DATA_BLOCK DB 1
VERSION : 0.1


  STRUCT
   STAT0 : CHAR ;
   STAT1 : CHAR ;
   STAT2 : CHAR ;
   STAT3 : CHAR ;
   STAT4 : CHAR ;
   STAT5 : CHAR ;
   STAT6 : CHAR ;
   STAT7 : CHAR ;
   STAT8 : CHAR ;
   STAT9 : CHAR ;
   STAT10 : CHAR ;
   STAT11 : CHAR ;
  END_STRUCT ;
BEGIN
   STAT0 := ' ';
   STAT1 := ' ';
   STAT2 := ' ';
   STAT3 := ' ';
   STAT4 := ' ';
   STAT5 := ' ';
   STAT6 := ' ';
   STAT7 := ' ';
   STAT8 := ' ';
   STAT9 := ' ';
   STAT10 := ' ';
   STAT11 := ' ';
END_DATA_BLOCK

DATA_BLOCK DB 2
VERSION : 0.1


  STRUCT
   STAT0 : CHAR ;
   STAT1 : CHAR ;
   STAT2 : CHAR ;
   STAT3 : CHAR ;
   STAT4 : CHAR ;
   STAT5 : CHAR ;
   STAT6 : CHAR ;
   STAT7 : CHAR ;
  END_STRUCT ;
BEGIN
   STAT0 := ' ';
   STAT1 := ' ';
   STAT2 := ' ';
   STAT3 := ' ';
   STAT4 := ' ';
   STAT5 := ' ';
   STAT6 := ' ';
   STAT7 := ' ';
END_DATA_BLOCK

DATA_BLOCK DB 3
VERSION : 0.1


  STRUCT
   STAT0 : INT ;
   STAT1 : BOOL ;
   STAT2 : INT ;
   STAT3 : BOOL ;
   STAT4 : BOOL ;
   STAT5 : BOOL ;
   STAT6 : BOOL ;
   STAT7 : BOOL ;
   STAT8 : BOOL ;
   STAT9 : BOOL ;
   STAT10 : BOOL ;
   STAT11 : BOOL ;
   STAT12 : BOOL ;
   STAT13 : BOOL ;
   STAT14 : BOOL ;
   STAT15 : INT ;
   STAT16 : INT ;
   STAT17 : INT ;
   STAT18 : INT ;
   STAT19 : CHAR  := '2';
   STAT20 : CHAR  := '8';
   STAT21 : INT ;
   STAT22 : CHAR  := '-';
   STAT23 : CHAR  := '-';
   STAT24 : CHAR  := '-';
   STAT25 : CHAR  := '-';
   STAT26 : CHAR  := '-';
   STAT27 : CHAR  := '-';
   STAT28 : CHAR  := '-';
   STAT29 : CHAR  := '-';
   STAT30 : CHAR  := '-';
   STAT31 : CHAR  := '-';
   STAT32 : CHAR  := '-';
   STAT33 : CHAR  := '-';
   STAT34 : CHAR  := '-';
   STAT35 : CHAR  := '-';
   STAT36 : CHAR  := '-';
   STAT37 : CHAR  := '-';
   STAT38 : CHAR  := '-';
   STAT39 : CHAR  := '-';
   STAT40 : CHAR  := '1';
   STAT41 : CHAR  := '2';
   STAT42 : CHAR  := '3';
   STAT43 : CHAR  := '4';
   STAT44 : CHAR  := '5';
   STAT45 : CHAR  := '6';
   STAT46 : CHAR  := '7';
   STAT47 : CHAR  := '8';
   STAT48 : CHAR  := '9';
   STAT49 : CHAR  := '0';
   STAT50 : INT ;
   STAT51 : INT ;
   STAT52 : INT ;
   STAT53 : INT ;
   STAT54 : INT ;
   STAT55 : CHAR  := '1';
   STAT56 : CHAR  := '4';
   STAT57 : CHAR  := '6';
   STAT58 : CHAR  := '1';
   STAT59 : CHAR  := '2';
   STAT60 : CHAR  := '3';
   STAT61 : CHAR  := '4';
   STAT62 : CHAR  := '5';
   STAT63 : CHAR  := '6';
   STAT64 : CHAR  := '7';
   STAT65 : CHAR  := '8';
   STAT66 : CHAR  := '9';
   STAT67 : CHAR  := '0';
   STAT68 : CHAR  := '1';
   STAT69 : CHAR  := '2';
   STAT70 : CHAR  := '3';
   STAT71 : CHAR  := '4';
   STAT72 : CHAR  := '5';
   STAT73 : CHAR  := '6';
   STAT74 : CHAR  := '7';
   STAT75 : CHAR  := '8';
   STAT76 : CHAR  := 'P';
   STAT77 : CHAR  := 'P';
   STAT78 : CHAR  := 'P';
   STAT79 : INT ;
   STAT80 : CHAR  := '0';
   STAT81 : CHAR  := '0';
   STAT82 : CHAR  := '0';
   STAT83 : CHAR  := '0';
   STAT84 : CHAR  := '0';
   STAT85 : CHAR  := '0';
   STAT86 : INT ;
   STAT87 : CHAR ;
   STAT88 : INT ;
   STAT89 : BOOL ;
   STAT90 : BOOL ;
   STAT91 : CHAR ;
   STAT92 : CHAR ;
   STAT93 : CHAR ;
   STAT94 : CHAR ;
   STAT95 : CHAR ;
   STAT96 : CHAR ;
   STAT97 : CHAR ;
   STAT98 : CHAR ;
   STAT99 : CHAR ;
   STAT100 : CHAR ;
   STAT101 : CHAR ;
   STAT102 : CHAR ;
   STAT103 : ARRAY  [1 .. 3 ] OF CHAR ;
   STAT104 : BOOL ;
   STAT105 : ARRAY  [1 .. 10 ] OF STRUCT
    STAT106 : REAL ;
    STAT107 : REAL ;
    STAT108 : REAL ;
   END_STRUCT ;
   STAT109 : CHAR ;
   STAT110 : CHAR ;
   STAT111 : ARRAY  [1 .. 10 ] OF REAL ;
   STAT112 : INT ;
   STAT113 : BOOL ;
   STAT114 : BOOL ;
   STAT115 : BOOL ;
  END_STRUCT ;
BEGIN
   STAT0 := 0;
   STAT1 := FALSE;
   STAT2 := 0;
   STAT3 := FALSE;
   STAT4 := FALSE;
   STAT5 := FALSE;
   STAT6 := FALSE;
   STAT7 := FALSE;
   STAT8 := FALSE;
   STAT9 := FALSE;
   STAT10 := FALSE;
   STAT11 := FALSE;
   STAT12 := FALSE;
   STAT13 := FALSE;
   STAT14 := FALSE;
   STAT15 := 0;
   STAT16 := 0;
   STAT17 := 0;
   STAT18 := 0;
   STAT19 := ' ';
   STAT20 := ' ';
   STAT21 := 0;
   STAT22 := '1';
   STAT23 := '2';
   STAT24 := '3';
   STAT25 := '4';
   STAT26 := '5';
   STAT27 := '$00';
   STAT28 := '7';
   STAT29 := '8';
   STAT30 := '9';
   STAT31 := '0';
   STAT32 := '1';
   STAT33 := '$00';
   STAT34 := '3';
   STAT35 := '4';
   STAT36 := '5';
   STAT37 := '6';
   STAT38 := '7';
   STAT39 := '$00';
   STAT40 := '-';
   STAT41 := '-';
   STAT42 := '-';
   STAT43 := '-';
   STAT44 := '-';
   STAT45 := '-';
   STAT46 := '-';
   STAT47 := '-';
   STAT48 := '-';
   STAT49 := '-';
   STAT50 := 0;
   STAT51 := 0;
   STAT52 := 0;
   STAT53 := 0;
   STAT54 := 0;
   STAT55 := '1';
   STAT56 := '2';
   STAT57 := '3';
   STAT58 := '$00';
   STAT59 := '$00';
   STAT60 := '$00';
   STAT61 := '$00';
   STAT62 := '$00';
   STAT63 := '$00';
   STAT64 := '$00';
   STAT65 := '$00';
   STAT66 := '$00';
   STAT67 := '$00';
   STAT68 := '$00';
   STAT69 := '$00';
   STAT70 := '$00';
   STAT71 := '$00';
   STAT72 := '$00';
   STAT73 := '$00';
   STAT74 := '$00';
   STAT75 := '$00';
   STAT76 := 'P';
   STAT77 := 'P';
   STAT78 := 'P';
   STAT79 := 0;
   STAT80 := '$00';
   STAT81 := '$00';
   STAT82 := '$00';
   STAT83 := '$00';
   STAT84 := '$00';
   STAT85 := '$00';
   STAT86 := 1;
   STAT87 := '1';
   STAT88 := 49;
   STAT89 := FALSE;
   STAT90 := FALSE;
   STAT91 := '-';
   STAT92 := '-';
   STAT93 := '-';
   STAT94 := '$00';
   STAT95 := '$00';
   STAT96 := '$00';
   STAT97 := '$00';
   STAT98 := '$00';
   STAT99 := '$00';
   STAT100 := '$00';
   STAT101 := '$00';
   STAT102 := '$00';
   STAT103[1] := '-';
   STAT103[2] := '-';
   STAT103[3] := '-';
   STAT104 := FALSE;
   STAT105[1].STAT106 := 1.616663e+004;
   STAT105[1].STAT107 := -7.696248e+003;
   STAT105[1].STAT108 := 1.325872e+004;
   STAT105[2].STAT106 := -8.515102e+003;
   STAT105[2].STAT107 := 3.194731e+000;
   STAT105[2].STAT108 := 2.146098e+004;
   STAT105[3].STAT106 := -3.152269e+003;
   STAT105[3].STAT107 := 5.230335e+001;
   STAT105[3].STAT108 := 1.702762e+004;
   STAT105[4].STAT106 := 4.876809e+003;
   STAT105[4].STAT107 := -1.412248e+003;
   STAT105[4].STAT108 := 3.514912e+004;
   STAT105[5].STAT106 := 0.000000e+000;
   STAT105[5].STAT107 := 0.000000e+000;
   STAT105[5].STAT108 := 0.000000e+000;
   STAT105[6].STAT106 := 0.000000e+000;
   STAT105[6].STAT107 := 0.000000e+000;
   STAT105[6].STAT108 := 0.000000e+000;
   STAT105[7].STAT106 := 0.000000e+000;
   STAT105[7].STAT107 := 0.000000e+000;
   STAT105[7].STAT108 := 0.000000e+000;
   STAT105[8].STAT106 := 0.000000e+000;
   STAT105[8].STAT107 := 0.000000e+000;
   STAT105[8].STAT108 := 0.000000e+000;
   STAT105[9].STAT106 := 0.000000e+000;
   STAT105[9].STAT107 := 0.000000e+000;
   STAT105[9].STAT108 := 0.000000e+000;
   STAT105[10].STAT106 := 0.000000e+000;
   STAT105[10].STAT107 := 0.000000e+000;
   STAT105[10].STAT108 := 0.000000e+000;
   STAT109 := '-';
   STAT110 := '-';
   STAT111[1] := -2.054582e+003;
   STAT111[2] := -2.149658e-001;
   STAT111[3] := -9.505859e+000;
   STAT111[4] := 1.638507e+003;
   STAT111[5] := 0.000000e+000;
   STAT111[6] := 0.000000e+000;
   STAT111[7] := 0.000000e+000;
   STAT111[8] := 0.000000e+000;
   STAT111[9] := 0.000000e+000;
   STAT111[10] := 0.000000e+000;
   STAT112 := 1;
   STAT113 := FALSE;
   STAT114 := FALSE;
   STAT115 := FALSE;
END_DATA_BLOCK

DATA_BLOCK DB 4
VERSION : 0.1


  STRUCT
   STAT0 : INT ;
   STAT1 : ARRAY  [1 .. 10 ] OF INT ;
   STAT2 : ARRAY  [1 .. 10 ] OF INT ;
   STAT3 : ARRAY  [1 .. 10 ] OF INT ;
  END_STRUCT ;
BEGIN
   STAT0 := 0;
   STAT1[1] := -32768;
   STAT1[2] := 17072;
   STAT1[3] := 17056;
   STAT1[4] := 16968;
   STAT1[5] := 0;
   STAT1[6] := 0;
   STAT1[7] := 0;
   STAT1[8] := 0;
   STAT1[9] := 0;
   STAT1[10] := 0;
   STAT2[1] := 5576;
   STAT2[2] := 1968;
   STAT2[3] := -1312;
   STAT2[4] := -1624;
   STAT2[5] := 0;
   STAT2[6] := 0;
   STAT2[7] := 0;
   STAT2[8] := 0;
   STAT2[9] := 0;
   STAT2[10] := 0;
   STAT3[1] := -1632;
   STAT3[2] := 13768;
   STAT3[3] := 27488;
   STAT3[4] := 27496;
   STAT3[5] := 0;
   STAT3[6] := 0;
   STAT3[7] := 0;
   STAT3[8] := 0;
   STAT3[9] := 0;
   STAT3[10] := 0;
END_DATA_BLOCK

DATA_BLOCK DB 5
VERSION : 0.1


  STRUCT
   STAT0 : INT ;
   STAT1 : ARRAY  [1 .. 10 ] OF BOOL ;
   STAT2 : ARRAY  [1 .. 10 ] OF BOOL ;
   STAT3 : BOOL ;
   STAT4 : BOOL ;
   STAT5 : BOOL ;
   STAT6 : ARRAY  [1 .. 10 ] OF BOOL ;
   STAT7 : ARRAY  [1 .. 10 ] OF BOOL ;
   STAT8 : ARRAY  [1 .. 10 ] OF INT  := 0;
   STAT9 : ARRAY  [1 .. 10 ] OF INT  := 0;
   STAT10 : ARRAY  [1 .. 10 ] OF INT  := 0;
   STAT11 : ARRAY  [1 .. 10 ] OF INT  := 0;
   STAT12 : ARRAY  [1 .. 10 ] OF INT  := 0;
   STAT13 : ARRAY  [1 .. 10 ] OF INT  := 0;
   STAT14 : ARRAY  [1 .. 10 ] OF INT  := 0;
   STAT15 : ARRAY  [1 .. 10 ] OF INT  := 0;
   STAT16 : ARRAY  [1 .. 10 ] OF INT  := 0;
   STAT17 : ARRAY  [1 .. 10 ] OF INT  := 0;
   STAT18 : ARRAY  [1 .. 10 ] OF BOOL ;
   STAT19 : ARRAY  [1 .. 10 ] OF BOOL ;
  END_STRUCT ;
BEGIN
   STAT0 := 0;
   STAT1[1] := FALSE;
   STAT1[2] := FALSE;
   STAT1[3] := FALSE;
   STAT1[4] := FALSE;
   STAT1[5] := FALSE;
   STAT1[6] := FALSE;
   STAT1[7] := FALSE;
   STAT1[8] := FALSE;
   STAT1[9] := FALSE;
   STAT1[10] := FALSE;
   STAT2[1] := FALSE;
   STAT2[2] := FALSE;
   STAT2[3] := FALSE;
   STAT2[4] := FALSE;
   STAT2[5] := FALSE;
   STAT2[6] := FALSE;
   STAT2[7] := FALSE;
   STAT2[8] := FALSE;
   STAT2[9] := FALSE;
   STAT2[10] := FALSE;
   STAT3 := FALSE;
   STAT4 := FALSE;
   STAT5 := FALSE;
   STAT6[1] := FALSE;
   STAT6[2] := FALSE;
   STAT6[3] := FALSE;
   STAT6[4] := FALSE;
   STAT6[5] := FALSE;
   STAT6[6] := FALSE;
   STAT6[7] := FALSE;
   STAT6[8] := FALSE;
   STAT6[9] := FALSE;
   STAT6[10] := FALSE;
   STAT7[1] := FALSE;
   STAT7[2] := FALSE;
   STAT7[3] := FALSE;
   STAT7[4] := FALSE;
   STAT7[5] := FALSE;
   STAT7[6] := FALSE;
   STAT7[7] := FALSE;
   STAT7[8] := FALSE;
   STAT7[9] := FALSE;
   STAT7[10] := FALSE;
   STAT8[1] := 0;
   STAT8[2] := 0;
   STAT8[3] := 0;
   STAT8[4] := 0;
   STAT8[5] := 0;
   STAT8[6] := 0;
   STAT8[7] := 0;
   STAT8[8] := 0;
   STAT8[9] := 0;
   STAT8[10] := 0;
   STAT9[1] := 0;
   STAT9[2] := 0;
   STAT9[3] := 0;
   STAT9[4] := 0;
   STAT9[5] := 0;
   STAT9[6] := 0;
   STAT9[7] := 0;
   STAT9[8] := 0;
   STAT9[9] := 0;
   STAT9[10] := 0;
   STAT10[1] := 0;
   STAT10[2] := 0;
   STAT10[3] := 0;
   STAT10[4] := 0;
   STAT10[5] := 0;
   STAT10[6] := 0;
   STAT10[7] := 0;
   STAT10[8] := 0;
   STAT10[9] := 0;
   STAT10[10] := 0;
   STAT11[1] := 0;
   STAT11[2] := 0;
   STAT11[3] := 0;
   STAT11[4] := 0;
   STAT11[5] := 0;
   STAT11[6] := 0;
   STAT11[7] := 0;
   STAT11[8] := 0;
   STAT11[9] := 0;
   STAT11[10] := 0;
   STAT12[1] := 0;
   STAT12[2] := 0;
   STAT12[3] := 0;
   STAT12[4] := 0;
   STAT12[5] := 0;
   STAT12[6] := 0;
   STAT12[7] := 0;
   STAT12[8] := 0;
   STAT12[9] := 0;
   STAT12[10] := 0;
   STAT13[1] := 0;
   STAT13[2] := 0;
   STAT13[3] := 0;
   STAT13[4] := 0;
   STAT13[5] := 0;
   STAT13[6] := 0;
   STAT13[7] := 0;
   STAT13[8] := 0;
   STAT13[9] := 0;
   STAT13[10] := 0;
   STAT14[1] := 0;
   STAT14[2] := 0;
   STAT14[3] := 0;
   STAT14[4] := 0;
   STAT14[5] := 0;
   STAT14[6] := 0;
   STAT14[7] := 0;
   STAT14[8] := 0;
   STAT14[9] := 0;
   STAT14[10] := 0;
   STAT15[1] := 0;
   STAT15[2] := 0;
   STAT15[3] := 0;
   STAT15[4] := 0;
   STAT15[5] := 0;
   STAT15[6] := 0;
   STAT15[7] := 0;
   STAT15[8] := 0;
   STAT15[9] := 0;
   STAT15[10] := 0;
   STAT16[1] := 0;
   STAT16[2] := 0;
   STAT16[3] := 0;
   STAT16[4] := 0;
   STAT16[5] := 0;
   STAT16[6] := 0;
   STAT16[7] := 0;
   STAT16[8] := 0;
   STAT16[9] := 0;
   STAT16[10] := 0;
   STAT17[1] := 0;
   STAT17[2] := 0;
   STAT17[3] := 0;
   STAT17[4] := 0;
   STAT17[5] := 0;
   STAT17[6] := 0;
   STAT17[7] := 0;
   STAT17[8] := 0;
   STAT17[9] := 0;
   STAT17[10] := 0;
   STAT18[1] := FALSE;
   STAT18[2] := FALSE;
   STAT18[3] := FALSE;
   STAT18[4] := FALSE;
   STAT18[5] := FALSE;
   STAT18[6] := FALSE;
   STAT18[7] := FALSE;
   STAT18[8] := FALSE;
   STAT18[9] := FALSE;
   STAT18[10] := FALSE;
   STAT19[1] := FALSE;
   STAT19[2] := FALSE;
   STAT19[3] := FALSE;
   STAT19[4] := FALSE;
   STAT19[5] := FALSE;
   STAT19[6] := FALSE;
   STAT19[7] := FALSE;
   STAT19[8] := FALSE;
   STAT19[9] := FALSE;
   STAT19[10] := FALSE;
END_DATA_BLOCK

DATA_BLOCK DB 6
VERSION : 0.0


  STRUCT
   STAT0 : BOOL ;
   STAT1 : BOOL ;
   STAT2 : BOOL ;
   STAT3 : BOOL ;
   STAT4 : BOOL ;
   STAT5 : BOOL ;
   STAT6 : BOOL ;
   STAT7 : BOOL ;
   STAT8 : BOOL ;
   STAT9 : BOOL ;
   STAT10 : BOOL ;
   STAT11 : BOOL ;
   STAT12 : BOOL ;
   STAT13 : S5TIME ;
   STAT14 : BOOL ;
   STAT15 : BOOL ;
   STAT16 : BOOL ;
   STAT17 : BOOL ;
   STAT18 : BOOL ;
   STAT19 : BOOL ;
   STAT20 : BOOL ;
   STAT21 : INT ;
  END_STRUCT ;
BEGIN
   STAT0 := FALSE;
   STAT1 := FALSE;
   STAT2 := FALSE;
   STAT3 := FALSE;
   STAT4 := FALSE;
   STAT5 := FALSE;
   STAT6 := FALSE;
   STAT7 := FALSE;
   STAT8 := FALSE;
   STAT9 := FALSE;
   STAT10 := TRUE;
   STAT11 := FALSE;
   STAT12 := TRUE;
   STAT13 := S5T#10S;
   STAT14 := FALSE;
   STAT15 := FALSE;
   STAT16 := FALSE;
   STAT17 := FALSE;
   STAT18 := FALSE;
   STAT19 := FALSE;
   STAT20 := TRUE;
   STAT21 := 4;
END_DATA_BLOCK

DATA_BLOCK DB 7
VERSION : 0.1


  STRUCT
   STAT0 : INT ;
   STAT1 : INT ;
   STAT2 : INT ;
   STAT3 : INT ;
   STAT4 : INT ;
   STAT5 : INT ;
   STAT6 : INT ;
   STAT7 : INT ;
   STAT8 : INT ;
   STAT9 : INT ;
   STAT10 : ARRAY  [1 .. 10 ] OF REAL ;
   STAT11 : ARRAY  [1 .. 10 ] OF REAL ;
   STAT12 : ARRAY  [1 .. 10 ] OF REAL ;
   STAT13 : ARRAY  [1 .. 10 ] OF REAL ;
   STAT14 : ARRAY  [1 .. 10 ] OF REAL ;
   STAT15 : ARRAY  [1 .. 10 ] OF INT  := 0;
   STAT16 : ARRAY  [1 .. 10 ] OF INT  := 0;
   STAT17 : ARRAY  [1 .. 10 ] OF INT  := 0;
   STAT18 : ARRAY  [1 .. 10 ] OF INT  := 0;
   STAT19 : ARRAY  [1 .. 10 ] OF INT  := 0;
   STAT20 : ARRAY  [1 .. 10 ] OF INT  := 0;
   STAT21 : ARRAY  [1 .. 10 ] OF INT  := 0;
   STAT22 : ARRAY  [1 .. 10 ] OF INT  := 0;
   STAT23 : ARRAY  [1 .. 10 ] OF INT  := 0;
   STAT24 : ARRAY  [1 .. 3 ] OF INT ;
   STAT25 : ARRAY  [1 .. 3 ] OF INT ;
   STAT26 : ARRAY  [1 .. 3 ] OF INT ;
   STAT27 : ARRAY  [1 .. 3 ] OF INT ;
   STAT28 : ARRAY  [1 .. 9 ] OF INT ;
   STAT29 : ARRAY  [1 .. 9 ] OF INT ;
   STAT30 : ARRAY  [1 .. 9 ] OF INT ;
   STAT31 : ARRAY  [1 .. 3 ] OF INT ;
   STAT32 : REAL ;
   STAT33 : REAL ;
   STAT34 : ARRAY  [1 .. 10 ] OF INT ;
   STAT35 : ARRAY  [1 .. 10 ] OF INT ;
   STAT36 : ARRAY  [1 .. 10 ] OF INT ;
   STAT37 : ARRAY  [1 .. 10 ] OF INT ;
   STAT38 : ARRAY  [1 .. 10 ] OF INT ;
   STAT39 : ARRAY  [1 .. 10 ] OF INT ;
   STAT40 : ARRAY  [1 .. 3 ] OF INT ;
   STAT41 : ARRAY  [1 .. 3 ] OF INT ;
   STAT42 : WORD ;
   STAT43 : ARRAY  [1 .. 10 ] OF REAL ;
   STAT44 : ARRAY  [1 .. 10 ] OF REAL ;
   STAT45 : ARRAY  [1 .. 10 ] OF REAL ;
  END_STRUCT ;
BEGIN
   STAT0 := 0;
   STAT1 := 0;
   STAT2 := 0;
   STAT3 := 0;
   STAT4 := 0;
   STAT5 := 0;
   STAT6 := 0;
   STAT7 := 0;
   STAT8 := 0;
   STAT9 := 0;
   STAT10[1] := -3.132816e+003;
   STAT10[2] := 2.383809e+004;
   STAT10[3] := 1.891266e+004;
   STAT10[4] := 1.#QNAN0e+000;
   STAT10[5] := 0.000000e+000;
   STAT10[6] := 0.000000e+000;
   STAT10[7] := 0.000000e+000;
   STAT10[8] := 0.000000e+000;
   STAT10[9] := 0.000000e+000;
   STAT10[10] := 0.000000e+000;
   STAT11[1] := 2.580549e+003;
   STAT11[2] := 4.758385e+003;
   STAT11[3] := 1.799429e+003;
   STAT11[4] := -3.709761e+003;
   STAT11[5] := 0.000000e+000;
   STAT11[6] := 0.000000e+000;
   STAT11[7] := 0.000000e+000;
   STAT11[8] := 0.000000e+000;
   STAT11[9] := 0.000000e+000;
   STAT11[10] := 0.000000e+000;
   STAT12[1] := 1.696806e+004;
   STAT12[2] := -5.077715e+003;
   STAT12[3] := -4.419669e+002;
   STAT12[4] := 2.768744e+003;
   STAT12[5] := 0.000000e+000;
   STAT12[6] := 0.000000e+000;
   STAT12[7] := 0.000000e+000;
   STAT12[8] := 0.000000e+000;
   STAT12[9] := 0.000000e+000;
   STAT12[10] := 0.000000e+000;
   STAT13[1] := 4.279937e+003;
   STAT13[2] := -3.930041e+003;
   STAT13[3] := 5.123809e+002;
   STAT13[4] := -1.760913e+004;
   STAT13[5] := 0.000000e+000;
   STAT13[6] := 0.000000e+000;
   STAT13[7] := 0.000000e+000;
   STAT13[8] := 0.000000e+000;
   STAT13[9] := 0.000000e+000;
   STAT13[10] := 0.000000e+000;
   STAT14[1] := 3.570063e+003;
   STAT14[2] := 1.178004e+004;
   STAT14[3] := 7.337619e+003;
   STAT14[4] := 2.545913e+004;
   STAT14[5] := 0.000000e+000;
   STAT14[6] := 0.000000e+000;
   STAT14[7] := 0.000000e+000;
   STAT14[8] := 0.000000e+000;
   STAT14[9] := 0.000000e+000;
   STAT14[10] := 0.000000e+000;
   STAT15[1] := 0;
   STAT15[2] := 0;
   STAT15[3] := 0;
   STAT15[4] := 0;
   STAT15[5] := 0;
   STAT15[6] := 0;
   STAT15[7] := 0;
   STAT15[8] := 0;
   STAT15[9] := 0;
   STAT15[10] := 0;
   STAT16[1] := 0;
   STAT16[2] := 0;
   STAT16[3] := 0;
   STAT16[4] := 0;
   STAT16[5] := 0;
   STAT16[6] := 0;
   STAT16[7] := 0;
   STAT16[8] := 0;
   STAT16[9] := 0;
   STAT16[10] := 0;
   STAT17[1] := 0;
   STAT17[2] := 0;
   STAT17[3] := 0;
   STAT17[4] := 0;
   STAT17[5] := 0;
   STAT17[6] := 0;
   STAT17[7] := 0;
   STAT17[8] := 0;
   STAT17[9] := 0;
   STAT17[10] := 0;
   STAT18[1] := 0;
   STAT18[2] := 0;
   STAT18[3] := 0;
   STAT18[4] := 0;
   STAT18[5] := 0;
   STAT18[6] := 0;
   STAT18[7] := 0;
   STAT18[8] := 0;
   STAT18[9] := 0;
   STAT18[10] := 0;
   STAT19[1] := 0;
   STAT19[2] := 0;
   STAT19[3] := 0;
   STAT19[4] := 0;
   STAT19[5] := 0;
   STAT19[6] := 0;
   STAT19[7] := 0;
   STAT19[8] := 0;
   STAT19[9] := 0;
   STAT19[10] := 0;
   STAT20[1] := 0;
   STAT20[2] := 0;
   STAT20[3] := 0;
   STAT20[4] := 0;
   STAT20[5] := 0;
   STAT20[6] := 0;
   STAT20[7] := 0;
   STAT20[8] := 0;
   STAT20[9] := 0;
   STAT20[10] := 0;
   STAT21[1] := 0;
   STAT21[2] := 0;
   STAT21[3] := 0;
   STAT21[4] := 0;
   STAT21[5] := 0;
   STAT21[6] := 0;
   STAT21[7] := 0;
   STAT21[8] := 0;
   STAT21[9] := 0;
   STAT21[10] := 0;
   STAT22[1] := 0;
   STAT22[2] := 0;
   STAT22[3] := 0;
   STAT22[4] := 0;
   STAT22[5] := 0;
   STAT22[6] := 0;
   STAT22[7] := 0;
   STAT22[8] := 0;
   STAT22[9] := 0;
   STAT22[10] := 0;
   STAT23[1] := 0;
   STAT23[2] := 0;
   STAT23[3] := 0;
   STAT23[4] := 0;
   STAT23[5] := 0;
   STAT23[6] := 0;
   STAT23[7] := 0;
   STAT23[8] := 0;
   STAT23[9] := 0;
   STAT23[10] := 0;
   STAT24[1] := 0;
   STAT24[2] := 0;
   STAT24[3] := 0;
   STAT25[1] := 0;
   STAT25[2] := 0;
   STAT25[3] := 0;
   STAT26[1] := 0;
   STAT26[2] := 0;
   STAT26[3] := 0;
   STAT27[1] := 51;
   STAT27[2] := 51;
   STAT27[3] := 51;
   STAT28[1] := 0;
   STAT28[2] := 0;
   STAT28[3] := 0;
   STAT28[4] := 0;
   STAT28[5] := 0;
   STAT28[6] := 0;
   STAT28[7] := 0;
   STAT28[8] := 0;
   STAT28[9] := 0;
   STAT29[1] := 0;
   STAT29[2] := 0;
   STAT29[3] := 0;
   STAT29[4] := 0;
   STAT29[5] := 0;
   STAT29[6] := 0;
   STAT29[7] := 0;
   STAT29[8] := 0;
   STAT29[9] := 0;
   STAT30[1] := 0;
   STAT30[2] := 0;
   STAT30[3] := 0;
   STAT30[4] := 0;
   STAT30[5] := 0;
   STAT30[6] := 0;
   STAT30[7] := 0;
   STAT30[8] := 0;
   STAT30[9] := 0;
   STAT31[1] := 49;
   STAT31[2] := 50;
   STAT31[3] := 51;
   STAT32 := 0.000000e+000;
   STAT33 := 0.000000e+000;
   STAT34[1] := 0;
   STAT34[2] := 0;
   STAT34[3] := 0;
   STAT34[4] := 0;
   STAT34[5] := 0;
   STAT34[6] := 0;
   STAT34[7] := 0;
   STAT34[8] := 0;
   STAT34[9] := 0;
   STAT34[10] := 0;
   STAT35[1] := 0;
   STAT35[2] := 0;
   STAT35[3] := 0;
   STAT35[4] := 0;
   STAT35[5] := 0;
   STAT35[6] := 0;
   STAT35[7] := 0;
   STAT35[8] := 0;
   STAT35[9] := 0;
   STAT35[10] := 0;
   STAT36[1] := 0;
   STAT36[2] := 0;
   STAT36[3] := 0;
   STAT36[4] := 0;
   STAT36[5] := 0;
   STAT36[6] := 0;
   STAT36[7] := 0;
   STAT36[8] := 0;
   STAT36[9] := 0;
   STAT36[10] := 0;
   STAT37[1] := 0;
   STAT37[2] := 0;
   STAT37[3] := 0;
   STAT37[4] := 0;
   STAT37[5] := 0;
   STAT37[6] := 0;
   STAT37[7] := 0;
   STAT37[8] := 0;
   STAT37[9] := 0;
   STAT37[10] := 0;
   STAT38[1] := 0;
   STAT38[2] := 0;
   STAT38[3] := 0;
   STAT38[4] := 0;
   STAT38[5] := 0;
   STAT38[6] := 0;
   STAT38[7] := 0;
   STAT38[8] := 0;
   STAT38[9] := 0;
   STAT38[10] := 0;
   STAT39[1] := 0;
   STAT39[2] := 0;
   STAT39[3] := 0;
   STAT39[4] := 0;
   STAT39[5] := 0;
   STAT39[6] := 0;
   STAT39[7] := 0;
   STAT39[8] := 0;
   STAT39[9] := 0;
   STAT39[10] := 0;
   STAT40[1] := 0;
   STAT40[2] := 0;
   STAT40[3] := 0;
   STAT41[1] := 0;
   STAT41[2] := 0;
   STAT41[3] := 0;
   STAT42 := W#16#96C7;
   STAT43[1] := 1.401610e+003;
   STAT43[2] := 5.370077e+003;
   STAT43[3] := 1.968209e+003;
   STAT43[4] := -4.097883e+003;
   STAT43[5] := 0.000000e+000;
   STAT43[6] := 0.000000e+000;
   STAT43[7] := 0.000000e+000;
   STAT43[8] := 0.000000e+000;
   STAT43[9] := 0.000000e+000;
   STAT43[10] := 0.000000e+000;
   STAT44[1] := 1.799841e+004;
   STAT44[2] := -5.547811e+003;
   STAT44[3] := -6.710018e+002;
   STAT44[4] := 3.114294e+003;
   STAT44[5] := 0.000000e+000;
   STAT44[6] := 0.000000e+000;
   STAT44[7] := 0.000000e+000;
   STAT44[8] := 0.000000e+000;
   STAT44[9] := 0.000000e+000;
   STAT44[10] := 0.000000e+000;
   STAT45[1] := -2.575992e+003;
   STAT45[2] := 2.431540e+004;
   STAT45[3] := 1.937619e+004;
   STAT45[4] := 1.#QNAN0e+000;
   STAT45[5] := 0.000000e+000;
   STAT45[6] := 0.000000e+000;
   STAT45[7] := 0.000000e+000;
   STAT45[8] := 0.000000e+000;
   STAT45[9] := 0.000000e+000;
   STAT45[10] := 0.000000e+000;
END_DATA_BLOCK

DATA_BLOCK DB 8
VERSION : 0.1


  STRUCT
   STAT0 : INT ;
   STAT1 : ARRAY  [1 .. 10 ] OF BOOL ;
   STAT2 : ARRAY  [1 .. 10 ] OF BOOL ;
  END_STRUCT ;
BEGIN
   STAT0 := 0;
   STAT1[1] := FALSE;
   STAT1[2] := FALSE;
   STAT1[3] := FALSE;
   STAT1[4] := FALSE;
   STAT1[5] := FALSE;
   STAT1[6] := FALSE;
   STAT1[7] := FALSE;
   STAT1[8] := FALSE;
   STAT1[9] := FALSE;
   STAT1[10] := FALSE;
   STAT2[1] := FALSE;
   STAT2[2] := FALSE;
   STAT2[3] := FALSE;
   STAT2[4] := FALSE;
   STAT2[5] := FALSE;
   STAT2[6] := FALSE;
   STAT2[7] := FALSE;
   STAT2[8] := FALSE;
   STAT2[9] := FALSE;
   STAT2[10] := FALSE;
END_DATA_BLOCK

DATA_BLOCK DB 9
VERSION : 0.0


  STRUCT
   STAT0 : ARRAY  [1 .. 10 ] OF REAL ;
   STAT1 : ARRAY  [1 .. 10 ] OF REAL ;
   STAT2 : ARRAY  [1 .. 10 ] OF BOOL ;
   STAT3 : ARRAY  [1 .. 10 ] OF BOOL ;
   STAT4 : ARRAY  [1 .. 10 ] OF BOOL ;
   STAT5 : ARRAY  [1 .. 10 ] OF BOOL ;
   STAT6 : BOOL ;
   STAT7 : ARRAY  [1 .. 10 ] OF BOOL  := FALSE;
  END_STRUCT ;
BEGIN
   STAT0[1] := 0.000000e+000;
   STAT0[2] := 0.000000e+000;
   STAT0[3] := 0.000000e+000;
   STAT0[4] := 0.000000e+000;
   STAT0[5] := 0.000000e+000;
   STAT0[6] := 0.000000e+000;
   STAT0[7] := 0.000000e+000;
   STAT0[8] := 0.000000e+000;
   STAT0[9] := 0.000000e+000;
   STAT0[10] := 0.000000e+000;
   STAT1[1] := 0.000000e+000;
   STAT1[2] := 0.000000e+000;
   STAT1[3] := 0.000000e+000;
   STAT1[4] := 0.000000e+000;
   STAT1[5] := 0.000000e+000;
   STAT1[6] := 0.000000e+000;
   STAT1[7] := 0.000000e+000;
   STAT1[8] := 0.000000e+000;
   STAT1[9] := 0.000000e+000;
   STAT1[10] := 0.000000e+000;
   STAT2[1] := FALSE;
   STAT2[2] := FALSE;
   STAT2[3] := FALSE;
   STAT2[4] := FALSE;
   STAT2[5] := FALSE;
   STAT2[6] := FALSE;
   STAT2[7] := FALSE;
   STAT2[8] := FALSE;
   STAT2[9] := FALSE;
   STAT2[10] := FALSE;
   STAT3[1] := FALSE;
   STAT3[2] := FALSE;
   STAT3[3] := FALSE;
   STAT3[4] := FALSE;
   STAT3[5] := FALSE;
   STAT3[6] := FALSE;
   STAT3[7] := FALSE;
   STAT3[8] := FALSE;
   STAT3[9] := FALSE;
   STAT3[10] := FALSE;
   STAT4[1] := FALSE;
   STAT4[2] := FALSE;
   STAT4[3] := FALSE;
   STAT4[4] := FALSE;
   STAT4[5] := FALSE;
   STAT4[6] := FALSE;
   STAT4[7] := FALSE;
   STAT4[8] := FALSE;
   STAT4[9] := FALSE;
   STAT4[10] := FALSE;
   STAT5[1] := FALSE;
   STAT5[2] := FALSE;
   STAT5[3] := FALSE;
   STAT5[4] := FALSE;
   STAT5[5] := FALSE;
   STAT5[6] := FALSE;
   STAT5[7] := FALSE;
   STAT5[8] := FALSE;
   STAT5[9] := FALSE;
   STAT5[10] := FALSE;
   STAT6 := FALSE;
   STAT7[1] := FALSE;
   STAT7[2] := FALSE;
   STAT7[3] := FALSE;
   STAT7[4] := FALSE;
   STAT7[5] := FALSE;
   STAT7[6] := FALSE;
   STAT7[7] := FALSE;
   STAT7[8] := FALSE;
   STAT7[9] := FALSE;
   STAT7[10] := FALSE;
END_DATA_BLOCK

DATA_BLOCK DB 10
VERSION : 0.1


  STRUCT
   STAT0 : INT ;
   STAT1 : REAL ;
   STAT2 : REAL  := 3.141593e+000;
   STAT3 : REAL ;
   STAT4 : REAL ;
   STAT5 : BOOL ;
  END_STRUCT ;
BEGIN
   STAT0 := 0;
   STAT1 := 0.000000e+000;
   STAT2 := 3.141593e+000;
   STAT3 := 0.000000e+000;
   STAT4 := 0.000000e+000;
   STAT5 := FALSE;
END_DATA_BLOCK

DATA_BLOCK DB 11
VERSION : 0.1


  STRUCT
   STAT0 : INT ;
   STAT1 : ARRAY  [1 .. 10 ] OF BOOL ;
  END_STRUCT ;
BEGIN
   STAT0 := 0;
   STAT1[1] := FALSE;
   STAT1[2] := FALSE;
   STAT1[3] := FALSE;
   STAT1[4] := FALSE;
   STAT1[5] := FALSE;
   STAT1[6] := FALSE;
   STAT1[7] := FALSE;
   STAT1[8] := FALSE;
   STAT1[9] := FALSE;
   STAT1[10] := FALSE;
END_DATA_BLOCK

DATA_BLOCK DB 12
VERSION : 0.1


  STRUCT
   STAT0 : INT ;
   STAT1 : REAL ;
   STAT2 : ARRAY  [1 .. 10 ] OF STRUCT
    STAT3 : REAL ;
    STAT4 : REAL ;
    STAT5 : REAL ;
   END_STRUCT ;
   STAT6 : ARRAY  [1 .. 10 ] OF REAL  := 0.000000e+000;
   STAT7 : ARRAY  [1 .. 10 ] OF BOOL ;
   STAT8 : REAL ;
   STAT9 : REAL ;
   STAT10 : REAL ;
   STAT11 : REAL ;
   STAT12 : ARRAY  [1 .. 10 ] OF REAL ;
   STAT13 : BOOL ;
  END_STRUCT ;
BEGIN
   STAT0 := 0;
   STAT1 := 5.000000e+000;
   STAT2[1].STAT3 := 0.000000e+000;
   STAT2[1].STAT4 := 0.000000e+000;
   STAT2[1].STAT5 := 0.000000e+000;
   STAT2[2].STAT3 := 0.000000e+000;
   STAT2[2].STAT4 := 0.000000e+000;
   STAT2[2].STAT5 := 0.000000e+000;
   STAT2[3].STAT3 := 0.000000e+000;
   STAT2[3].STAT4 := 0.000000e+000;
   STAT2[3].STAT5 := 0.000000e+000;
   STAT2[4].STAT3 := 0.000000e+000;
   STAT2[4].STAT4 := 0.000000e+000;
   STAT2[4].STAT5 := 0.000000e+000;
   STAT2[5].STAT3 := 0.000000e+000;
   STAT2[5].STAT4 := 0.000000e+000;
   STAT2[5].STAT5 := 0.000000e+000;
   STAT2[6].STAT3 := 0.000000e+000;
   STAT2[6].STAT4 := 0.000000e+000;
   STAT2[6].STAT5 := 0.000000e+000;
   STAT2[7].STAT3 := 0.000000e+000;
   STAT2[7].STAT4 := 0.000000e+000;
   STAT2[7].STAT5 := 0.000000e+000;
   STAT2[8].STAT3 := 0.000000e+000;
   STAT2[8].STAT4 := 0.000000e+000;
   STAT2[8].STAT5 := 0.000000e+000;
   STAT2[9].STAT3 := 0.000000e+000;
   STAT2[9].STAT4 := 0.000000e+000;
   STAT2[9].STAT5 := 0.000000e+000;
   STAT2[10].STAT3 := 0.000000e+000;
   STAT2[10].STAT4 := 0.000000e+000;
   STAT2[10].STAT5 := 0.000000e+000;
   STAT6[1] := 1.623795e+004;
   STAT6[2] := 1.623795e+004;
   STAT6[3] := 1.623795e+004;
   STAT6[4] := 1.623795e+004;
   STAT6[5] := 0.000000e+000;
   STAT6[6] := 0.000000e+000;
   STAT6[7] := 0.000000e+000;
   STAT6[8] := 0.000000e+000;
   STAT6[9] := 0.000000e+000;
   STAT6[10] := 0.000000e+000;
   STAT7[1] := FALSE;
   STAT7[2] := FALSE;
   STAT7[3] := FALSE;
   STAT7[4] := FALSE;
   STAT7[5] := FALSE;
   STAT7[6] := FALSE;
   STAT7[7] := FALSE;
   STAT7[8] := FALSE;
   STAT7[9] := FALSE;
   STAT7[10] := FALSE;
   STAT8 := 0.000000e+000;
   STAT9 := 0.000000e+000;
   STAT10 := 0.000000e+000;
   STAT11 := 0.000000e+000;
   STAT12[1] := 1.577482e+004;
   STAT12[2] := 1.577482e+004;
   STAT12[3] := 1.577482e+004;
   STAT12[4] := 1.577482e+004;
   STAT12[5] := 0.000000e+000;
   STAT12[6] := 0.000000e+000;
   STAT12[7] := 0.000000e+000;
   STAT12[8] := 0.000000e+000;
   STAT12[9] := 0.000000e+000;
   STAT12[10] := 0.000000e+000;
   STAT13 := FALSE;
END_DATA_BLOCK

DATA_BLOCK DB 13
VERSION : 0.1


  STRUCT
   STAT0 : INT ;
   STAT1 : BOOL ;
   STAT2 : BOOL ;
   STAT3 : BOOL ;
   STAT4 : ARRAY  [1 .. 10 ] OF BOOL ;
   STAT5 : ARRAY  [1 .. 10 ] OF BOOL ;
   STAT6 : ARRAY  [1 .. 10 ] OF WORD ;
   STAT7 : ARRAY  [1 .. 10 ] OF WORD ;
   STAT8 : ARRAY  [1 .. 10 ] OF WORD ;
   STAT9 : BOOL ;
   STAT10 : BOOL ;
   STAT11 : BOOL ;
   STAT12 : BOOL ;
   STAT13 : ARRAY  [1 .. 10 ] OF BOOL ;
   STAT14 : ARRAY  [1 .. 10 ] OF BOOL ;
   STAT15 : BOOL ;
   STAT16 : BOOL ;
   STAT17 : BOOL ;
   STAT18 : ARRAY  [1 .. 10 ] OF BOOL ;
  END_STRUCT ;
BEGIN
   STAT0 := 0;
   STAT1 := FALSE;
   STAT2 := FALSE;
   STAT3 := FALSE;
   STAT4[1] := FALSE;
   STAT4[2] := FALSE;
   STAT4[3] := FALSE;
   STAT4[4] := FALSE;
   STAT4[5] := FALSE;
   STAT4[6] := FALSE;
   STAT4[7] := FALSE;
   STAT4[8] := FALSE;
   STAT4[9] := FALSE;
   STAT4[10] := FALSE;
   STAT5[1] := FALSE;
   STAT5[2] := FALSE;
   STAT5[3] := FALSE;
   STAT5[4] := FALSE;
   STAT5[5] := FALSE;
   STAT5[6] := FALSE;
   STAT5[7] := FALSE;
   STAT5[8] := FALSE;
   STAT5[9] := FALSE;
   STAT5[10] := FALSE;
   STAT6[1] := W#16#0;
   STAT6[2] := W#16#0;
   STAT6[3] := W#16#0;
   STAT6[4] := W#16#0;
   STAT6[5] := W#16#0;
   STAT6[6] := W#16#0;
   STAT6[7] := W#16#0;
   STAT6[8] := W#16#0;
   STAT6[9] := W#16#0;
   STAT6[10] := W#16#0;
   STAT7[1] := W#16#0;
   STAT7[2] := W#16#0;
   STAT7[3] := W#16#0;
   STAT7[4] := W#16#0;
   STAT7[5] := W#16#0;
   STAT7[6] := W#16#0;
   STAT7[7] := W#16#0;
   STAT7[8] := W#16#0;
   STAT7[9] := W#16#0;
   STAT7[10] := W#16#0;
   STAT8[1] := W#16#0;
   STAT8[2] := W#16#0;
   STAT8[3] := W#16#0;
   STAT8[4] := W#16#0;
   STAT8[5] := W#16#0;
   STAT8[6] := W#16#0;
   STAT8[7] := W#16#0;
   STAT8[8] := W#16#0;
   STAT8[9] := W#16#0;
   STAT8[10] := W#16#0;
   STAT9 := FALSE;
   STAT10 := FALSE;
   STAT11 := FALSE;
   STAT12 := FALSE;
   STAT13[1] := FALSE;
   STAT13[2] := FALSE;
   STAT13[3] := FALSE;
   STAT13[4] := FALSE;
   STAT13[5] := FALSE;
   STAT13[6] := FALSE;
   STAT13[7] := FALSE;
   STAT13[8] := FALSE;
   STAT13[9] := FALSE;
   STAT13[10] := FALSE;
   STAT14[1] := FALSE;
   STAT14[2] := FALSE;
   STAT14[3] := FALSE;
   STAT14[4] := FALSE;
   STAT14[5] := FALSE;
   STAT14[6] := FALSE;
   STAT14[7] := FALSE;
   STAT14[8] := FALSE;
   STAT14[9] := FALSE;
   STAT14[10] := FALSE;
   STAT15 := FALSE;
   STAT16 := FALSE;
   STAT17 := FALSE;
   STAT18[1] := FALSE;
   STAT18[2] := FALSE;
   STAT18[3] := FALSE;
   STAT18[4] := FALSE;
   STAT18[5] := FALSE;
   STAT18[6] := FALSE;
   STAT18[7] := FALSE;
   STAT18[8] := FALSE;
   STAT18[9] := FALSE;
   STAT18[10] := FALSE;
END_DATA_BLOCK

DATA_BLOCK DB 14
VERSION : 0.1


  STRUCT
   STAT0 : INT ;
   STAT1 : BOOL ;
   STAT2 : INT ;
   STAT3 : INT ;
   STAT4 : INT ;
   STAT5 : BYTE ;
   STAT6 : REAL ;
   STAT7 : REAL ;
   STAT8 : REAL ;
   STAT9 : ARRAY  [1 .. 10 ] OF STRUCT
    STAT10 : REAL ;
    STAT11 : REAL ;
    STAT12 : REAL ;
   END_STRUCT ;
   STAT13 : BYTE ;
   STAT14 : BOOL ;
   STAT15 : BOOL ;
  END_STRUCT ;
BEGIN
   STAT0 := 0;
   STAT1 := FALSE;
   STAT2 := 0;
   STAT3 := 0;
   STAT4 := 0;
   STAT5 := B#16#0;
   STAT6 := 0.000000e+000;
   STAT7 := 0.000000e+000;
   STAT8 := 0.000000e+000;
   STAT9[1].STAT10 := -1.247000e+003;
   STAT9[1].STAT11 := -2.249000e+003;
   STAT9[1].STAT12 := -1.848000e+003;
   STAT9[2].STAT10 := -1.272000e+003;
   STAT9[2].STAT11 := -1.746000e+003;
   STAT9[2].STAT12 := -1.743000e+003;
   STAT9[3].STAT10 := -1.267000e+003;
   STAT9[3].STAT11 := -9.240000e+002;
   STAT9[3].STAT12 := -3.489000e+003;
   STAT9[4].STAT10 := -1.256000e+003;
   STAT9[4].STAT11 := -2.183000e+003;
   STAT9[4].STAT12 := -1.842000e+003;
   STAT9[5].STAT10 := 0.000000e+000;
   STAT9[5].STAT11 := 0.000000e+000;
   STAT9[5].STAT12 := 0.000000e+000;
   STAT9[6].STAT10 := 0.000000e+000;
   STAT9[6].STAT11 := 0.000000e+000;
   STAT9[6].STAT12 := 0.000000e+000;
   STAT9[7].STAT10 := 0.000000e+000;
   STAT9[7].STAT11 := 0.000000e+000;
   STAT9[7].STAT12 := 0.000000e+000;
   STAT9[8].STAT10 := 0.000000e+000;
   STAT9[8].STAT11 := 0.000000e+000;
   STAT9[8].STAT12 := 0.000000e+000;
   STAT9[9].STAT10 := 0.000000e+000;
   STAT9[9].STAT11 := 0.000000e+000;
   STAT9[9].STAT12 := 0.000000e+000;
   STAT9[10].STAT10 := 0.000000e+000;
   STAT9[10].STAT11 := 0.000000e+000;
   STAT9[10].STAT12 := 0.000000e+000;
   STAT13 := B#16#0;
   STAT14 := FALSE;
   STAT15 := FALSE;
END_DATA_BLOCK

DATA_BLOCK DB 15
VERSION : 0.0


  STRUCT
   STAT0 : INT ;
   STAT1 : INT ;
   STAT2 : INT ;
   STAT3 : INT ;
   STAT4 : ARRAY  [1 .. 15 ] OF INT ;
   STAT5 : ARRAY  [1 .. 15 ] OF INT ;
   STAT6 : ARRAY  [1 .. 15 ] OF INT ;
   STAT7 : ARRAY  [1 .. 15 ] OF BOOL ;
  END_STRUCT ;
BEGIN
   STAT0 := 0;
   STAT1 := 0;
   STAT2 := 0;
   STAT3 := 0;
   STAT4[1] := 0;
   STAT4[2] := 0;
   STAT4[3] := 0;
   STAT4[4] := 0;
   STAT4[5] := 0;
   STAT4[6] := 0;
   STAT4[7] := 0;
   STAT4[8] := 0;
   STAT4[9] := 0;
   STAT4[10] := 0;
   STAT4[11] := 0;
   STAT4[12] := 0;
   STAT4[13] := 0;
   STAT4[14] := 0;
   STAT4[15] := 0;
   STAT5[1] := 0;
   STAT5[2] := 0;
   STAT5[3] := 0;
   STAT5[4] := 0;
   STAT5[5] := 0;
   STAT5[6] := 0;
   STAT5[7] := 0;
   STAT5[8] := 0;
   STAT5[9] := 0;
   STAT5[10] := 0;
   STAT5[11] := 0;
   STAT5[12] := 0;
   STAT5[13] := 0;
   STAT5[14] := 0;
   STAT5[15] := 0;
   STAT6[1] := 0;
   STAT6[2] := 0;
   STAT6[3] := 0;
   STAT6[4] := 0;
   STAT6[5] := 0;
   STAT6[6] := 0;
   STAT6[7] := 0;
   STAT6[8] := 0;
   STAT6[9] := 0;
   STAT6[10] := 0;
   STAT6[11] := 0;
   STAT6[12] := 0;
   STAT6[13] := 0;
   STAT6[14] := 0;
   STAT6[15] := 0;
   STAT7[1] := FALSE;
   STAT7[2] := FALSE;
   STAT7[3] := FALSE;
   STAT7[4] := FALSE;
   STAT7[5] := FALSE;
   STAT7[6] := FALSE;
   STAT7[7] := FALSE;
   STAT7[8] := FALSE;
   STAT7[9] := FALSE;
   STAT7[10] := FALSE;
   STAT7[11] := FALSE;
   STAT7[12] := FALSE;
   STAT7[13] := FALSE;
   STAT7[14] := FALSE;
   STAT7[15] := FALSE;
END_DATA_BLOCK

DATA_BLOCK DB 16
VERSION : 0.1


  STRUCT
   STAT0 : INT ;
   STAT1 : ARRAY  [1 .. 10 ] OF BOOL  := FALSE;
  END_STRUCT ;
BEGIN
   STAT0 := 0;
   STAT1[1] := FALSE;
   STAT1[2] := FALSE;
   STAT1[3] := FALSE;
   STAT1[4] := FALSE;
   STAT1[5] := FALSE;
   STAT1[6] := FALSE;
   STAT1[7] := FALSE;
   STAT1[8] := FALSE;
   STAT1[9] := FALSE;
   STAT1[10] := FALSE;
END_DATA_BLOCK

DATA_BLOCK DB 17
VERSION : 0.1


  STRUCT
   STAT0 : INT ;
   STAT1 : BOOL ;
  END_STRUCT ;
BEGIN
   STAT0 := 0;
   STAT1 := FALSE;
END_DATA_BLOCK

DATA_BLOCK DB 18
VERSION : 0.1


  STRUCT
   STAT0 : BYTE ;
   STAT1 : INT ;
   STAT2 : WORD ;
   STAT3 : INT ;
   STAT4 : INT ;
   STAT5 : INT ;
   STAT6 : INT ;
   STAT7 : INT ;
  END_STRUCT ;
BEGIN
   STAT0 := B#16#4;
   STAT1 := -67;
   STAT2 := W#16#FFBD;
   STAT3 := 3;
   STAT4 := 3;
   STAT5 := 3;
   STAT6 := 3;
   STAT7 := 3;
END_DATA_BLOCK

DATA_BLOCK DB 19
VERSION : 0.1


  STRUCT
   STAT0 : BOOL ;
   STAT1 : BOOL ;
   STAT2 : BOOL ;
   STAT3 : BOOL ;
   STAT4 : BOOL ;
   STAT5 : BOOL ;
   STAT6 : BOOL ;
   STAT7 : BOOL ;
   STAT8 : BOOL ;
   STAT9 : BOOL ;
   STAT10 : BOOL ;
   STAT11 : BOOL ;
   STAT12 : BOOL ;
   STAT13 : BOOL ;
   STAT14 : BOOL ;
   STAT15 : BOOL ;
   STAT16 : BOOL ;
   STAT17 : BOOL ;
   STAT18 : BOOL ;
   STAT19 : BOOL ;
   STAT20 : BOOL ;
   STAT21 : BOOL ;
   STAT22 : BOOL ;
   STAT23 : BOOL ;
   STAT24 : BOOL ;
   STAT25 : BOOL ;
   STAT26 : BOOL ;
   STAT27 : BOOL ;
   STAT28 : BOOL ;
   STAT29 : BOOL ;
   STAT30 : BOOL ;
   STAT31 : BOOL ;
  END_STRUCT ;
BEGIN
   STAT0 := FALSE;
   STAT1 := FALSE;
   STAT2 := FALSE;
   STAT3 := FALSE;
   STAT4 := FALSE;
   STAT5 := FALSE;
   STAT6 := FALSE;
   STAT7 := FALSE;
   STAT8 := FALSE;
   STAT9 := FALSE;
   STAT10 := FALSE;
   STAT11 := FALSE;
   STAT12 := FALSE;
   STAT13 := FALSE;
   STAT14 := FALSE;
   STAT15 := FALSE;
   STAT16 := FALSE;
   STAT17 := FALSE;
   STAT18 := FALSE;
   STAT19 := FALSE;
   STAT20 := FALSE;
   STAT21 := FALSE;
   STAT22 := FALSE;
   STAT23 := FALSE;
   STAT24 := FALSE;
   STAT25 := FALSE;
   STAT26 := FALSE;
   STAT27 := FALSE;
   STAT28 := FALSE;
   STAT29 := FALSE;
   STAT30 := FALSE;
   STAT31 := FALSE;
END_DATA_BLOCK

DATA_BLOCK DB 20
VERSION : 0.1


  STRUCT
   STAT0 : ARRAY  [1 .. 10 ] OF STRUCT
    STAT1 : REAL ;
    STAT2 : REAL ;
    STAT3 : REAL ;
   END_STRUCT ;
   STAT4 : INT ;
  END_STRUCT ;
BEGIN
   STAT0[1].STAT1 := -5.394847e+003;
   STAT0[1].STAT2 := -1.542576e+003;
   STAT0[1].STAT3 := -2.054582e+003;
   STAT0[2].STAT1 := 8.890132e+002;
   STAT0[2].STAT2 := -1.497894e+003;
   STAT0[2].STAT3 := -2.149658e-001;
   STAT0[3].STAT1 := 8.919878e+002;
   STAT0[3].STAT2 := -1.090076e+003;
   STAT0[3].STAT3 := -9.505859e+000;
   STAT0[4].STAT1 := 8.918486e+002;
   STAT0[4].STAT2 := -2.388537e+003;
   STAT0[4].STAT3 := 1.638507e+003;
   STAT0[5].STAT1 := 0.000000e+000;
   STAT0[5].STAT2 := 0.000000e+000;
   STAT0[5].STAT3 := 0.000000e+000;
   STAT0[6].STAT1 := 0.000000e+000;
   STAT0[6].STAT2 := 0.000000e+000;
   STAT0[6].STAT3 := 0.000000e+000;
   STAT0[7].STAT1 := 0.000000e+000;
   STAT0[7].STAT2 := 0.000000e+000;
   STAT0[7].STAT3 := 0.000000e+000;
   STAT0[8].STAT1 := 0.000000e+000;
   STAT0[8].STAT2 := 0.000000e+000;
   STAT0[8].STAT3 := 0.000000e+000;
   STAT0[9].STAT1 := 0.000000e+000;
   STAT0[9].STAT2 := 0.000000e+000;
   STAT0[9].STAT3 := 0.000000e+000;
   STAT0[10].STAT1 := 0.000000e+000;
   STAT0[10].STAT2 := 0.000000e+000;
   STAT0[10].STAT3 := 0.000000e+000;
   STAT4 := 30;
END_DATA_BLOCK

DATA_BLOCK DB 21
VERSION : 0.1


  STRUCT
   STAT0 : INT ;
   STAT1 : INT ;
   STAT2 : INT ;
  END_STRUCT ;
BEGIN
   STAT0 := 1;
   STAT1 := -109;
   STAT2 := 89;
END_DATA_BLOCK

DATA_BLOCK DB 22
VERSION : 0.0


  STRUCT
   STAT0 : ARRAY  [1 .. 10 ] OF REAL ;
   STAT1 : ARRAY  [1 .. 10 ] OF REAL ;
   STAT2 : ARRAY  [1 .. 10 ] OF REAL ;
   STAT3 : ARRAY  [1 .. 10 ] OF STRUCT
    STAT4 : REAL ;
    STAT5 : REAL ;
    STAT6 : REAL ;
   END_STRUCT ;
   STAT7 : ARRAY  [1 .. 10 ] OF STRUCT
    STAT8 : REAL ;
    STAT9 : REAL ;
    STAT10 : REAL ;
   END_STRUCT ;
   STAT11 : ARRAY  [1 .. 10 ] OF STRUCT
    STAT12 : REAL ;
    STAT13 : REAL ;
    STAT14 : REAL ;
   END_STRUCT ;
   STAT15 : ARRAY  [1 .. 10 ] OF STRUCT
    STAT16 : REAL ;
    STAT17 : REAL ;
    STAT18 : REAL ;
   END_STRUCT ;
   STAT19 : ARRAY  [1 .. 10 ] OF STRUCT
    STAT20 : REAL ;
    STAT21 : REAL ;
    STAT22 : REAL ;
   END_STRUCT ;
   STAT23 : ARRAY  [1 .. 10, 1 .. 10 ] OF STRUCT
    STAT24 : REAL ;
    STAT25 : REAL ;
    STAT26 : REAL ;
   END_STRUCT ;
   STAT27 : ARRAY  [1 .. 10 ] OF BOOL ;
   STAT28 : ARRAY  [1 .. 10, 1 .. 10, 1 .. 10 ] OF REAL ;
   STAT29 : ARRAY  [1 .. 10, 1 .. 10 ] OF STRUCT
    STAT30 : REAL ;
    STAT31 : REAL ;
    STAT32 : REAL ;
   END_STRUCT ;
   STAT33 : ARRAY  [1 .. 10, 1 .. 10, 1 .. 10 ] OF REAL ;
   STAT34 : ARRAY  [1 .. 10 ] OF INT ;
   STAT35 : ARRAY  [1 .. 10 ] OF BOOL ;
   STAT36 : ARRAY  [1 .. 10 ] OF BOOL ;
   STAT37 : ARRAY  [1 .. 10 ] OF BOOL ;
   STAT38 : ARRAY  [1 .. 10 ] OF STRUCT
    STAT39 : REAL ;
    STAT40 : REAL ;
    STAT41 : REAL ;
   END_STRUCT ;
   STAT42 : ARRAY  [1 .. 10 ] OF STRUCT
    STAT43 : REAL ;
    STAT44 : REAL ;
    STAT45 : REAL ;
   END_STRUCT ;
   STAT46 : INT ;
   STAT47 : INT ;
   STAT48 : ARRAY  [1 .. 10 ] OF STRUCT
    STAT49 : REAL ;
    STAT50 : REAL ;
    STAT51 : REAL ;
   END_STRUCT ;
   STAT52 : ARRAY  [1 .. 10 ] OF STRUCT
    STAT53 : REAL ;
    STAT54 : REAL ;
    STAT55 : REAL ;
   END_STRUCT ;
   STAT56 : INT ;
   STAT57 : ARRAY  [1 .. 10 ] OF STRUCT
    STAT58 : REAL ;
    STAT59 : REAL ;
    STAT60 : REAL ;
   END_STRUCT ;
   STAT61 : REAL ;
   STAT62 : REAL ;
   STAT63 : REAL ;
   STAT64 : ARRAY  [1 .. 10 ] OF STRUCT
    STAT65 : REAL ;
    STAT66 : REAL ;
    STAT67 : REAL ;
   END_STRUCT ;
   STAT68 : BOOL  := TRUE;
   STAT69 : BOOL ;
   STAT70 : BOOL ;
   STAT71 : ARRAY  [1 .. 10 ] OF BOOL ;
  END_STRUCT ;
BEGIN
   STAT0[1] := 7.058228e+002;
   STAT0[2] := 2.481013e+002;
   STAT0[3] := -1.660759e+002;
   STAT0[4] := -2.055696e+002;
   STAT0[5] := 0.000000e+000;
   STAT0[6] := 0.000000e+000;
   STAT0[7] := 0.000000e+000;
   STAT0[8] := 0.000000e+000;
   STAT0[9] := 0.000000e+000;
   STAT0[10] := 0.000000e+000;
   STAT1[1] := -4.147848e+003;
   STAT1[2] := 2.161013e+003;
   STAT1[3] := 2.158987e+003;
   STAT1[4] := 2.147848e+003;
   STAT1[5] := 0.000000e+000;
   STAT1[6] := 0.000000e+000;
   STAT1[7] := 0.000000e+000;
   STAT1[8] := 0.000000e+000;
   STAT1[9] := 0.000000e+000;
   STAT1[10] := 0.000000e+000;
   STAT2[1] := -2.065823e+002;
   STAT2[2] := 1.742785e+003;
   STAT2[3] := 3.479494e+003;
   STAT2[4] := 3.480506e+003;
   STAT2[5] := 0.000000e+000;
   STAT2[6] := 0.000000e+000;
   STAT2[7] := 0.000000e+000;
   STAT2[8] := 0.000000e+000;
   STAT2[9] := 0.000000e+000;
   STAT2[10] := 0.000000e+000;
   STAT3[1].STAT4 := 0.000000e+000;
   STAT3[1].STAT5 := 0.000000e+000;
   STAT3[1].STAT6 := 0.000000e+000;
   STAT3[2].STAT4 := 0.000000e+000;
   STAT3[2].STAT5 := 0.000000e+000;
   STAT3[2].STAT6 := 0.000000e+000;
   STAT3[3].STAT4 := 0.000000e+000;
   STAT3[3].STAT5 := 0.000000e+000;
   STAT3[3].STAT6 := 0.000000e+000;
   STAT3[4].STAT4 := 0.000000e+000;
   STAT3[4].STAT5 := 0.000000e+000;
   STAT3[4].STAT6 := 0.000000e+000;
   STAT3[5].STAT4 := 0.000000e+000;
   STAT3[5].STAT5 := 0.000000e+000;
   STAT3[5].STAT6 := 0.000000e+000;
   STAT3[6].STAT4 := 0.000000e+000;
   STAT3[6].STAT5 := 0.000000e+000;
   STAT3[6].STAT6 := 0.000000e+000;
   STAT3[7].STAT4 := 0.000000e+000;
   STAT3[7].STAT5 := 0.000000e+000;
   STAT3[7].STAT6 := 0.000000e+000;
   STAT3[8].STAT4 := 0.000000e+000;
   STAT3[8].STAT5 := 0.000000e+000;
   STAT3[8].STAT6 := 0.000000e+000;
   STAT3[9].STAT4 := 0.000000e+000;
   STAT3[9].STAT5 := 0.000000e+000;
   STAT3[9].STAT6 := 0.000000e+000;
   STAT3[10].STAT4 := 0.000000e+000;
   STAT3[10].STAT5 := 0.000000e+000;
   STAT3[10].STAT6 := 0.000000e+000;
   STAT7[1].STAT8 := 0.000000e+000;
   STAT7[1].STAT9 := 0.000000e+000;
   STAT7[1].STAT10 := 0.000000e+000;
   STAT7[2].STAT8 := 0.000000e+000;
   STAT7[2].STAT9 := 0.000000e+000;
   STAT7[2].STAT10 := 0.000000e+000;
   STAT7[3].STAT8 := 0.000000e+000;
   STAT7[3].STAT9 := 0.000000e+000;
   STAT7[3].STAT10 := 0.000000e+000;
   STAT7[4].STAT8 := 0.000000e+000;
   STAT7[4].STAT9 := 0.000000e+000;
   STAT7[4].STAT10 := 0.000000e+000;
   STAT7[5].STAT8 := 0.000000e+000;
   STAT7[5].STAT9 := 0.000000e+000;
   STAT7[5].STAT10 := 0.000000e+000;
   STAT7[6].STAT8 := 0.000000e+000;
   STAT7[6].STAT9 := 0.000000e+000;
   STAT7[6].STAT10 := 0.000000e+000;
   STAT7[7].STAT8 := 0.000000e+000;
   STAT7[7].STAT9 := 0.000000e+000;
   STAT7[7].STAT10 := 0.000000e+000;
   STAT7[8].STAT8 := 0.000000e+000;
   STAT7[8].STAT9 := 0.000000e+000;
   STAT7[8].STAT10 := 0.000000e+000;
   STAT7[9].STAT8 := 0.000000e+000;
   STAT7[9].STAT9 := 0.000000e+000;
   STAT7[9].STAT10 := 0.000000e+000;
   STAT7[10].STAT8 := 0.000000e+000;
   STAT7[10].STAT9 := 0.000000e+000;
   STAT7[10].STAT10 := 0.000000e+000;
   STAT11[1].STAT12 := 1.692603e+004;
   STAT11[1].STAT13 := -7.793991e+003;
   STAT11[1].STAT14 := 1.076110e+004;
   STAT11[2].STAT12 := -7.713949e+003;
   STAT11[2].STAT13 := 2.731981e+002;
   STAT11[2].STAT14 := 1.898631e+004;
   STAT11[3].STAT12 := -2.346739e+003;
   STAT11[3].STAT13 := -2.176596e+002;
   STAT11[3].STAT14 := 1.453762e+004;
   STAT11[4].STAT12 := 5.915027e+003;
   STAT11[4].STAT13 := -6.246460e+002;
   STAT11[4].STAT14 := 3.265903e+004;
   STAT11[5].STAT12 := 0.000000e+000;
   STAT11[5].STAT13 := 0.000000e+000;
   STAT11[5].STAT14 := 0.000000e+000;
   STAT11[6].STAT12 := 0.000000e+000;
   STAT11[6].STAT13 := 0.000000e+000;
   STAT11[6].STAT14 := 0.000000e+000;
   STAT11[7].STAT12 := 0.000000e+000;
   STAT11[7].STAT13 := 0.000000e+000;
   STAT11[7].STAT14 := 0.000000e+000;
   STAT11[8].STAT12 := 0.000000e+000;
   STAT11[8].STAT13 := 0.000000e+000;
   STAT11[8].STAT14 := 0.000000e+000;
   STAT11[9].STAT12 := 0.000000e+000;
   STAT11[9].STAT13 := 0.000000e+000;
   STAT11[9].STAT14 := 0.000000e+000;
   STAT11[10].STAT12 := 0.000000e+000;
   STAT11[10].STAT13 := 0.000000e+000;
   STAT11[10].STAT14 := 0.000000e+000;
   STAT15[1].STAT16 := 0.000000e+000;
   STAT15[1].STAT17 := 0.000000e+000;
   STAT15[1].STAT18 := 0.000000e+000;
   STAT15[2].STAT16 := 0.000000e+000;
   STAT15[2].STAT17 := 0.000000e+000;
   STAT15[2].STAT18 := 0.000000e+000;
   STAT15[3].STAT16 := 0.000000e+000;
   STAT15[3].STAT17 := 0.000000e+000;
   STAT15[3].STAT18 := 0.000000e+000;
   STAT15[4].STAT16 := 0.000000e+000;
   STAT15[4].STAT17 := 0.000000e+000;
   STAT15[4].STAT18 := 0.000000e+000;
   STAT15[5].STAT16 := 0.000000e+000;
   STAT15[5].STAT17 := 0.000000e+000;
   STAT15[5].STAT18 := 0.000000e+000;
   STAT15[6].STAT16 := 0.000000e+000;
   STAT15[6].STAT17 := 0.000000e+000;
   STAT15[6].STAT18 := 0.000000e+000;
   STAT15[7].STAT16 := 0.000000e+000;
   STAT15[7].STAT17 := 0.000000e+000;
   STAT15[7].STAT18 := 0.000000e+000;
   STAT15[8].STAT16 := 0.000000e+000;
   STAT15[8].STAT17 := 0.000000e+000;
   STAT15[8].STAT18 := 0.000000e+000;
   STAT15[9].STAT16 := 0.000000e+000;
   STAT15[9].STAT17 := 0.000000e+000;
   STAT15[9].STAT18 := 0.000000e+000;
   STAT15[10].STAT16 := 0.000000e+000;
   STAT15[10].STAT17 := 0.000000e+000;
   STAT15[10].STAT18 := 0.000000e+000;
   STAT19[1].STAT20 := 1.035156e-002;
   STAT19[1].STAT21 := 1.989746e-003;
   STAT19[1].STAT22 := 2.144531e-002;
   STAT19[2].STAT20 := -2.441406e-006;
   STAT19[2].STAT21 := -9.918213e-005;
   STAT19[2].STAT22 := 0.000000e+000;
   STAT19[3].STAT20 := -1.674316e-002;
   STAT19[3].STAT21 := 2.777100e-004;
   STAT19[3].STAT22 := 5.878906e-003;
   STAT19[4].STAT20 := 0.000000e+000;
   STAT19[4].STAT21 := 0.000000e+000;
   STAT19[4].STAT22 := 0.000000e+000;
   STAT19[5].STAT20 := 0.000000e+000;
   STAT19[5].STAT21 := 0.000000e+000;
   STAT19[5].STAT22 := 0.000000e+000;
   STAT19[6].STAT20 := 0.000000e+000;
   STAT19[6].STAT21 := 0.000000e+000;
   STAT19[6].STAT22 := 0.000000e+000;
   STAT19[7].STAT20 := 0.000000e+000;
   STAT19[7].STAT21 := 0.000000e+000;
   STAT19[7].STAT22 := 0.000000e+000;
   STAT19[8].STAT20 := 0.000000e+000;
   STAT19[8].STAT21 := 0.000000e+000;
   STAT19[8].STAT22 := 0.000000e+000;
   STAT19[9].STAT20 := 0.000000e+000;
   STAT19[9].STAT21 := 0.000000e+000;
   STAT19[9].STAT22 := 0.000000e+000;
   STAT19[10].STAT20 := 0.000000e+000;
   STAT19[10].STAT21 := 0.000000e+000;
   STAT19[10].STAT22 := 0.000000e+000;
   STAT23[1, 1].STAT24 := 0.000000e+000;
   STAT23[1, 1].STAT25 := 0.000000e+000;
   STAT23[1, 1].STAT26 := 0.000000e+000;
   STAT23[1, 2].STAT24 := 0.000000e+000;
   STAT23[1, 2].STAT25 := 0.000000e+000;
   STAT23[1, 2].STAT26 := 0.000000e+000;
   STAT23[1, 3].STAT24 := 0.000000e+000;
   STAT23[1, 3].STAT25 := 0.000000e+000;
   STAT23[1, 3].STAT26 := 0.000000e+000;
   STAT23[1, 4].STAT24 := 0.000000e+000;
   STAT23[1, 4].STAT25 := 0.000000e+000;
   STAT23[1, 4].STAT26 := 0.000000e+000;
   STAT23[1, 5].STAT24 := 0.000000e+000;
   STAT23[1, 5].STAT25 := 0.000000e+000;
   STAT23[1, 5].STAT26 := 0.000000e+000;
   STAT23[1, 6].STAT24 := 0.000000e+000;
   STAT23[1, 6].STAT25 := 0.000000e+000;
   STAT23[1, 6].STAT26 := 0.000000e+000;
   STAT23[1, 7].STAT24 := 0.000000e+000;
   STAT23[1, 7].STAT25 := 0.000000e+000;
   STAT23[1, 7].STAT26 := 0.000000e+000;
   STAT23[1, 8].STAT24 := 0.000000e+000;
   STAT23[1, 8].STAT25 := 0.000000e+000;
   STAT23[1, 8].STAT26 := 0.000000e+000;
   STAT23[1, 9].STAT24 := 0.000000e+000;
   STAT23[1, 9].STAT25 := 0.000000e+000;
   STAT23[1, 9].STAT26 := 0.000000e+000;
   STAT23[1, 10].STAT24 := 0.000000e+000;
   STAT23[1, 10].STAT25 := 0.000000e+000;
   STAT23[1, 10].STAT26 := 0.000000e+000;
   STAT23[2, 1].STAT24 := 0.000000e+000;
   STAT23[2, 1].STAT25 := 0.000000e+000;
   STAT23[2, 1].STAT26 := 0.000000e+000;
   STAT23[2, 2].STAT24 := 0.000000e+000;
   STAT23[2, 2].STAT25 := 0.000000e+000;
   STAT23[2, 2].STAT26 := 0.000000e+000;
   STAT23[2, 3].STAT24 := 0.000000e+000;
   STAT23[2, 3].STAT25 := 0.000000e+000;
   STAT23[2, 3].STAT26 := 0.000000e+000;
   STAT23[2, 4].STAT24 := 0.000000e+000;
   STAT23[2, 4].STAT25 := 0.000000e+000;
   STAT23[2, 4].STAT26 := 0.000000e+000;
   STAT23[2, 5].STAT24 := 0.000000e+000;
   STAT23[2, 5].STAT25 := 0.000000e+000;
   STAT23[2, 5].STAT26 := 0.000000e+000;
   STAT23[2, 6].STAT24 := 0.000000e+000;
   STAT23[2, 6].STAT25 := 0.000000e+000;
   STAT23[2, 6].STAT26 := 0.000000e+000;
   STAT23[2, 7].STAT24 := 0.000000e+000;
   STAT23[2, 7].STAT25 := 0.000000e+000;
   STAT23[2, 7].STAT26 := 0.000000e+000;
   STAT23[2, 8].STAT24 := 0.000000e+000;
   STAT23[2, 8].STAT25 := 0.000000e+000;
   STAT23[2, 8].STAT26 := 0.000000e+000;
   STAT23[2, 9].STAT24 := 0.000000e+000;
   STAT23[2, 9].STAT25 := 0.000000e+000;
   STAT23[2, 9].STAT26 := 0.000000e+000;
   STAT23[2, 10].STAT24 := 0.000000e+000;
   STAT23[2, 10].STAT25 := 0.000000e+000;
   STAT23[2, 10].STAT26 := 0.000000e+000;
   STAT23[3, 1].STAT24 := 0.000000e+000;
   STAT23[3, 1].STAT25 := 0.000000e+000;
   STAT23[3, 1].STAT26 := 0.000000e+000;
   STAT23[3, 2].STAT24 := 0.000000e+000;
   STAT23[3, 2].STAT25 := 0.000000e+000;
   STAT23[3, 2].STAT26 := 0.000000e+000;
   STAT23[3, 3].STAT24 := 0.000000e+000;
   STAT23[3, 3].STAT25 := 0.000000e+000;
   STAT23[3, 3].STAT26 := 0.000000e+000;
   STAT23[3, 4].STAT24 := 0.000000e+000;
   STAT23[3, 4].STAT25 := 0.000000e+000;
   STAT23[3, 4].STAT26 := 0.000000e+000;
   STAT23[3, 5].STAT24 := 0.000000e+000;
   STAT23[3, 5].STAT25 := 0.000000e+000;
   STAT23[3, 5].STAT26 := 0.000000e+000;
   STAT23[3, 6].STAT24 := 0.000000e+000;
   STAT23[3, 6].STAT25 := 0.000000e+000;
   STAT23[3, 6].STAT26 := 0.000000e+000;
   STAT23[3, 7].STAT24 := 0.000000e+000;
   STAT23[3, 7].STAT25 := 0.000000e+000;
   STAT23[3, 7].STAT26 := 0.000000e+000;
   STAT23[3, 8].STAT24 := 0.000000e+000;
   STAT23[3, 8].STAT25 := 0.000000e+000;
   STAT23[3, 8].STAT26 := 0.000000e+000;
   STAT23[3, 9].STAT24 := 0.000000e+000;
   STAT23[3, 9].STAT25 := 0.000000e+000;
   STAT23[3, 9].STAT26 := 0.000000e+000;
   STAT23[3, 10].STAT24 := 0.000000e+000;
   STAT23[3, 10].STAT25 := 0.000000e+000;
   STAT23[3, 10].STAT26 := 0.000000e+000;
   STAT23[4, 1].STAT24 := 0.000000e+000;
   STAT23[4, 1].STAT25 := 0.000000e+000;
   STAT23[4, 1].STAT26 := 0.000000e+000;
   STAT23[4, 2].STAT24 := 0.000000e+000;
   STAT23[4, 2].STAT25 := 0.000000e+000;
   STAT23[4, 2].STAT26 := 0.000000e+000;
   STAT23[4, 3].STAT24 := 0.000000e+000;
   STAT23[4, 3].STAT25 := 0.000000e+000;
   STAT23[4, 3].STAT26 := 0.000000e+000;
   STAT23[4, 4].STAT24 := 0.000000e+000;
   STAT23[4, 4].STAT25 := 0.000000e+000;
   STAT23[4, 4].STAT26 := 0.000000e+000;
   STAT23[4, 5].STAT24 := 0.000000e+000;
   STAT23[4, 5].STAT25 := 0.000000e+000;
   STAT23[4, 5].STAT26 := 0.000000e+000;
   STAT23[4, 6].STAT24 := 0.000000e+000;
   STAT23[4, 6].STAT25 := 0.000000e+000;
   STAT23[4, 6].STAT26 := 0.000000e+000;
   STAT23[4, 7].STAT24 := 0.000000e+000;
   STAT23[4, 7].STAT25 := 0.000000e+000;
   STAT23[4, 7].STAT26 := 0.000000e+000;
   STAT23[4, 8].STAT24 := 0.000000e+000;
   STAT23[4, 8].STAT25 := 0.000000e+000;
   STAT23[4, 8].STAT26 := 0.000000e+000;
   STAT23[4, 9].STAT24 := 0.000000e+000;
   STAT23[4, 9].STAT25 := 0.000000e+000;
   STAT23[4, 9].STAT26 := 0.000000e+000;
   STAT23[4, 10].STAT24 := 0.000000e+000;
   STAT23[4, 10].STAT25 := 0.000000e+000;
   STAT23[4, 10].STAT26 := 0.000000e+000;
   STAT23[5, 1].STAT24 := 0.000000e+000;
   STAT23[5, 1].STAT25 := 0.000000e+000;
   STAT23[5, 1].STAT26 := 0.000000e+000;
   STAT23[5, 2].STAT24 := 0.000000e+000;
   STAT23[5, 2].STAT25 := 0.000000e+000;
   STAT23[5, 2].STAT26 := 0.000000e+000;
   STAT23[5, 3].STAT24 := 0.000000e+000;
   STAT23[5, 3].STAT25 := 0.000000e+000;
   STAT23[5, 3].STAT26 := 0.000000e+000;
   STAT23[5, 4].STAT24 := 0.000000e+000;
   STAT23[5, 4].STAT25 := 0.000000e+000;
   STAT23[5, 4].STAT26 := 0.000000e+000;
   STAT23[5, 5].STAT24 := 0.000000e+000;
   STAT23[5, 5].STAT25 := 0.000000e+000;
   STAT23[5, 5].STAT26 := 0.000000e+000;
   STAT23[5, 6].STAT24 := 0.000000e+000;
   STAT23[5, 6].STAT25 := 0.000000e+000;
   STAT23[5, 6].STAT26 := 0.000000e+000;
   STAT23[5, 7].STAT24 := 0.000000e+000;
   STAT23[5, 7].STAT25 := 0.000000e+000;
   STAT23[5, 7].STAT26 := 0.000000e+000;
   STAT23[5, 8].STAT24 := 0.000000e+000;
   STAT23[5, 8].STAT25 := 0.000000e+000;
   STAT23[5, 8].STAT26 := 0.000000e+000;
   STAT23[5, 9].STAT24 := 0.000000e+000;
   STAT23[5, 9].STAT25 := 0.000000e+000;
   STAT23[5, 9].STAT26 := 0.000000e+000;
   STAT23[5, 10].STAT24 := 0.000000e+000;
   STAT23[5, 10].STAT25 := 0.000000e+000;
   STAT23[5, 10].STAT26 := 0.000000e+000;
   STAT23[6, 1].STAT24 := 0.000000e+000;
   STAT23[6, 1].STAT25 := 0.000000e+000;
   STAT23[6, 1].STAT26 := 0.000000e+000;
   STAT23[6, 2].STAT24 := 0.000000e+000;
   STAT23[6, 2].STAT25 := 0.000000e+000;
   STAT23[6, 2].STAT26 := 0.000000e+000;
   STAT23[6, 3].STAT24 := 0.000000e+000;
   STAT23[6, 3].STAT25 := 0.000000e+000;
   STAT23[6, 3].STAT26 := 0.000000e+000;
   STAT23[6, 4].STAT24 := 0.000000e+000;
   STAT23[6, 4].STAT25 := 0.000000e+000;
   STAT23[6, 4].STAT26 := 0.000000e+000;
   STAT23[6, 5].STAT24 := 0.000000e+000;
   STAT23[6, 5].STAT25 := 0.000000e+000;
   STAT23[6, 5].STAT26 := 0.000000e+000;
   STAT23[6, 6].STAT24 := 0.000000e+000;
   STAT23[6, 6].STAT25 := 0.000000e+000;
   STAT23[6, 6].STAT26 := 0.000000e+000;
   STAT23[6, 7].STAT24 := 0.000000e+000;
   STAT23[6, 7].STAT25 := 0.000000e+000;
   STAT23[6, 7].STAT26 := 0.000000e+000;
   STAT23[6, 8].STAT24 := 0.000000e+000;
   STAT23[6, 8].STAT25 := 0.000000e+000;
   STAT23[6, 8].STAT26 := 0.000000e+000;
   STAT23[6, 9].STAT24 := 0.000000e+000;
   STAT23[6, 9].STAT25 := 0.000000e+000;
   STAT23[6, 9].STAT26 := 0.000000e+000;
   STAT23[6, 10].STAT24 := 0.000000e+000;
   STAT23[6, 10].STAT25 := 0.000000e+000;
   STAT23[6, 10].STAT26 := 0.000000e+000;
   STAT23[7, 1].STAT24 := 0.000000e+000;
   STAT23[7, 1].STAT25 := 0.000000e+000;
   STAT23[7, 1].STAT26 := 0.000000e+000;
   STAT23[7, 2].STAT24 := 0.000000e+000;
   STAT23[7, 2].STAT25 := 0.000000e+000;
   STAT23[7, 2].STAT26 := 0.000000e+000;
   STAT23[7, 3].STAT24 := 0.000000e+000;
   STAT23[7, 3].STAT25 := 0.000000e+000;
   STAT23[7, 3].STAT26 := 0.000000e+000;
   STAT23[7, 4].STAT24 := 0.000000e+000;
   STAT23[7, 4].STAT25 := 0.000000e+000;
   STAT23[7, 4].STAT26 := 0.000000e+000;
   STAT23[7, 5].STAT24 := 0.000000e+000;
   STAT23[7, 5].STAT25 := 0.000000e+000;
   STAT23[7, 5].STAT26 := 0.000000e+000;
   STAT23[7, 6].STAT24 := 0.000000e+000;
   STAT23[7, 6].STAT25 := 0.000000e+000;
   STAT23[7, 6].STAT26 := 0.000000e+000;
   STAT23[7, 7].STAT24 := 0.000000e+000;
   STAT23[7, 7].STAT25 := 0.000000e+000;
   STAT23[7, 7].STAT26 := 0.000000e+000;
   STAT23[7, 8].STAT24 := 0.000000e+000;
   STAT23[7, 8].STAT25 := 0.000000e+000;
   STAT23[7, 8].STAT26 := 0.000000e+000;
   STAT23[7, 9].STAT24 := 0.000000e+000;
   STAT23[7, 9].STAT25 := 0.000000e+000;
   STAT23[7, 9].STAT26 := 0.000000e+000;
   STAT23[7, 10].STAT24 := 0.000000e+000;
   STAT23[7, 10].STAT25 := 0.000000e+000;
   STAT23[7, 10].STAT26 := 0.000000e+000;
   STAT23[8, 1].STAT24 := 0.000000e+000;
   STAT23[8, 1].STAT25 := 0.000000e+000;
   STAT23[8, 1].STAT26 := 0.000000e+000;
   STAT23[8, 2].STAT24 := 0.000000e+000;
   STAT23[8, 2].STAT25 := 0.000000e+000;
   STAT23[8, 2].STAT26 := 0.000000e+000;
   STAT23[8, 3].STAT24 := 0.000000e+000;
   STAT23[8, 3].STAT25 := 0.000000e+000;
   STAT23[8, 3].STAT26 := 0.000000e+000;
   STAT23[8, 4].STAT24 := 0.000000e+000;
   STAT23[8, 4].STAT25 := 0.000000e+000;
   STAT23[8, 4].STAT26 := 0.000000e+000;
   STAT23[8, 5].STAT24 := 0.000000e+000;
   STAT23[8, 5].STAT25 := 0.000000e+000;
   STAT23[8, 5].STAT26 := 0.000000e+000;
   STAT23[8, 6].STAT24 := 0.000000e+000;
   STAT23[8, 6].STAT25 := 0.000000e+000;
   STAT23[8, 6].STAT26 := 0.000000e+000;
   STAT23[8, 7].STAT24 := 0.000000e+000;
   STAT23[8, 7].STAT25 := 0.000000e+000;
   STAT23[8, 7].STAT26 := 0.000000e+000;
   STAT23[8, 8].STAT24 := 0.000000e+000;
   STAT23[8, 8].STAT25 := 0.000000e+000;
   STAT23[8, 8].STAT26 := 0.000000e+000;
   STAT23[8, 9].STAT24 := 0.000000e+000;
   STAT23[8, 9].STAT25 := 0.000000e+000;
   STAT23[8, 9].STAT26 := 0.000000e+000;
   STAT23[8, 10].STAT24 := 0.000000e+000;
   STAT23[8, 10].STAT25 := 0.000000e+000;
   STAT23[8, 10].STAT26 := 0.000000e+000;
   STAT23[9, 1].STAT24 := 0.000000e+000;
   STAT23[9, 1].STAT25 := 0.000000e+000;
   STAT23[9, 1].STAT26 := 0.000000e+000;
   STAT23[9, 2].STAT24 := 0.000000e+000;
   STAT23[9, 2].STAT25 := 0.000000e+000;
   STAT23[9, 2].STAT26 := 0.000000e+000;
   STAT23[9, 3].STAT24 := 0.000000e+000;
   STAT23[9, 3].STAT25 := 0.000000e+000;
   STAT23[9, 3].STAT26 := 0.000000e+000;
   STAT23[9, 4].STAT24 := 0.000000e+000;
   STAT23[9, 4].STAT25 := 0.000000e+000;
   STAT23[9, 4].STAT26 := 0.000000e+000;
   STAT23[9, 5].STAT24 := 0.000000e+000;
   STAT23[9, 5].STAT25 := 0.000000e+000;
   STAT23[9, 5].STAT26 := 0.000000e+000;
   STAT23[9, 6].STAT24 := 0.000000e+000;
   STAT23[9, 6].STAT25 := 0.000000e+000;
   STAT23[9, 6].STAT26 := 0.000000e+000;
   STAT23[9, 7].STAT24 := 0.000000e+000;
   STAT23[9, 7].STAT25 := 0.000000e+000;
   STAT23[9, 7].STAT26 := 0.000000e+000;
   STAT23[9, 8].STAT24 := 0.000000e+000;
   STAT23[9, 8].STAT25 := 0.000000e+000;
   STAT23[9, 8].STAT26 := 0.000000e+000;
   STAT23[9, 9].STAT24 := 0.000000e+000;
   STAT23[9, 9].STAT25 := 0.000000e+000;
   STAT23[9, 9].STAT26 := 0.000000e+000;
   STAT23[9, 10].STAT24 := 0.000000e+000;
   STAT23[9, 10].STAT25 := 0.000000e+000;
   STAT23[9, 10].STAT26 := 0.000000e+000;
   STAT23[10, 1].STAT24 := 0.000000e+000;
   STAT23[10, 1].STAT25 := 0.000000e+000;
   STAT23[10, 1].STAT26 := 0.000000e+000;
   STAT23[10, 2].STAT24 := 0.000000e+000;
   STAT23[10, 2].STAT25 := 0.000000e+000;
   STAT23[10, 2].STAT26 := 0.000000e+000;
   STAT23[10, 3].STAT24 := 0.000000e+000;
   STAT23[10, 3].STAT25 := 0.000000e+000;
   STAT23[10, 3].STAT26 := 0.000000e+000;
   STAT23[10, 4].STAT24 := 0.000000e+000;
   STAT23[10, 4].STAT25 := 0.000000e+000;
   STAT23[10, 4].STAT26 := 0.000000e+000;
   STAT23[10, 5].STAT24 := 0.000000e+000;
   STAT23[10, 5].STAT25 := 0.000000e+000;
   STAT23[10, 5].STAT26 := 0.000000e+000;
   STAT23[10, 6].STAT24 := 0.000000e+000;
   STAT23[10, 6].STAT25 := 0.000000e+000;
   STAT23[10, 6].STAT26 := 0.000000e+000;
   STAT23[10, 7].STAT24 := 0.000000e+000;
   STAT23[10, 7].STAT25 := 0.000000e+000;
   STAT23[10, 7].STAT26 := 0.000000e+000;
   STAT23[10, 8].STAT24 := 0.000000e+000;
   STAT23[10, 8].STAT25 := 0.000000e+000;
   STAT23[10, 8].STAT26 := 0.000000e+000;
   STAT23[10, 9].STAT24 := 0.000000e+000;
   STAT23[10, 9].STAT25 := 0.000000e+000;
   STAT23[10, 9].STAT26 := 0.000000e+000;
   STAT23[10, 10].STAT24 := 0.000000e+000;
   STAT23[10, 10].STAT25 := 0.000000e+000;
   STAT23[10, 10].STAT26 := 0.000000e+000;
   STAT27[1] := FALSE;
   STAT27[2] := FALSE;
   STAT27[3] := FALSE;
   STAT27[4] := FALSE;
   STAT27[5] := FALSE;
   STAT27[6] := FALSE;
   STAT27[7] := FALSE;
   STAT27[8] := FALSE;
   STAT27[9] := FALSE;
   STAT27[10] := FALSE;
   STAT28[1, 1, 1] := 0.000000e+000;
   STAT28[1, 1, 2] := 0.000000e+000;
   STAT28[1, 1, 3] := 0.000000e+000;
   STAT28[1, 1, 4] := 0.000000e+000;
   STAT28[1, 1, 5] := 0.000000e+000;
   STAT28[1, 1, 6] := 0.000000e+000;
   STAT28[1, 1, 7] := 0.000000e+000;
   STAT28[1, 1, 8] := 0.000000e+000;
   STAT28[1, 1, 9] := 0.000000e+000;
   STAT28[1, 1, 10] := 0.000000e+000;
   STAT28[1, 2, 1] := 0.000000e+000;
   STAT28[1, 2, 2] := 0.000000e+000;
   STAT28[1, 2, 3] := 0.000000e+000;
   STAT28[1, 2, 4] := 0.000000e+000;
   STAT28[1, 2, 5] := 0.000000e+000;
   STAT28[1, 2, 6] := 0.000000e+000;
   STAT28[1, 2, 7] := 0.000000e+000;
   STAT28[1, 2, 8] := 0.000000e+000;
   STAT28[1, 2, 9] := 0.000000e+000;
   STAT28[1, 2, 10] := 0.000000e+000;
   STAT28[1, 3, 1] := 0.000000e+000;
   STAT28[1, 3, 2] := 0.000000e+000;
   STAT28[1, 3, 3] := 0.000000e+000;
   STAT28[1, 3, 4] := 0.000000e+000;
   STAT28[1, 3, 5] := 0.000000e+000;
   STAT28[1, 3, 6] := 0.000000e+000;
   STAT28[1, 3, 7] := 0.000000e+000;
   STAT28[1, 3, 8] := 0.000000e+000;
   STAT28[1, 3, 9] := 0.000000e+000;
   STAT28[1, 3, 10] := 0.000000e+000;
   STAT28[1, 4, 1] := 0.000000e+000;
   STAT28[1, 4, 2] := 0.000000e+000;
   STAT28[1, 4, 3] := 0.000000e+000;
   STAT28[1, 4, 4] := 0.000000e+000;
   STAT28[1, 4, 5] := 0.000000e+000;
   STAT28[1, 4, 6] := 0.000000e+000;
   STAT28[1, 4, 7] := 0.000000e+000;
   STAT28[1, 4, 8] := 0.000000e+000;
   STAT28[1, 4, 9] := 0.000000e+000;
   STAT28[1, 4, 10] := 0.000000e+000;
   STAT28[1, 5, 1] := 0.000000e+000;
   STAT28[1, 5, 2] := 0.000000e+000;
   STAT28[1, 5, 3] := 0.000000e+000;
   STAT28[1, 5, 4] := 0.000000e+000;
   STAT28[1, 5, 5] := 0.000000e+000;
   STAT28[1, 5, 6] := 0.000000e+000;
   STAT28[1, 5, 7] := 0.000000e+000;
   STAT28[1, 5, 8] := 0.000000e+000;
   STAT28[1, 5, 9] := 0.000000e+000;
   STAT28[1, 5, 10] := 0.000000e+000;
   STAT28[1, 6, 1] := 0.000000e+000;
   STAT28[1, 6, 2] := 0.000000e+000;
   STAT28[1, 6, 3] := 0.000000e+000;
   STAT28[1, 6, 4] := 0.000000e+000;
   STAT28[1, 6, 5] := 0.000000e+000;
   STAT28[1, 6, 6] := 0.000000e+000;
   STAT28[1, 6, 7] := 0.000000e+000;
   STAT28[1, 6, 8] := 0.000000e+000;
   STAT28[1, 6, 9] := 0.000000e+000;
   STAT28[1, 6, 10] := 0.000000e+000;
   STAT28[1, 7, 1] := 0.000000e+000;
   STAT28[1, 7, 2] := 0.000000e+000;
   STAT28[1, 7, 3] := 0.000000e+000;
   STAT28[1, 7, 4] := 0.000000e+000;
   STAT28[1, 7, 5] := 0.000000e+000;
   STAT28[1, 7, 6] := 0.000000e+000;
   STAT28[1, 7, 7] := 0.000000e+000;
   STAT28[1, 7, 8] := 0.000000e+000;
   STAT28[1, 7, 9] := 0.000000e+000;
   STAT28[1, 7, 10] := 0.000000e+000;
   STAT28[1, 8, 1] := 0.000000e+000;
   STAT28[1, 8, 2] := 0.000000e+000;
   STAT28[1, 8, 3] := 0.000000e+000;
   STAT28[1, 8, 4] := 0.000000e+000;
   STAT28[1, 8, 5] := 0.000000e+000;
   STAT28[1, 8, 6] := 0.000000e+000;
   STAT28[1, 8, 7] := 0.000000e+000;
   STAT28[1, 8, 8] := 0.000000e+000;
   STAT28[1, 8, 9] := 0.000000e+000;
   STAT28[1, 8, 10] := 0.000000e+000;
   STAT28[1, 9, 1] := 0.000000e+000;
   STAT28[1, 9, 2] := 0.000000e+000;
   STAT28[1, 9, 3] := 0.000000e+000;
   STAT28[1, 9, 4] := 0.000000e+000;
   STAT28[1, 9, 5] := 0.000000e+000;
   STAT28[1, 9, 6] := 0.000000e+000;
   STAT28[1, 9, 7] := 0.000000e+000;
   STAT28[1, 9, 8] := 0.000000e+000;
   STAT28[1, 9, 9] := 0.000000e+000;
   STAT28[1, 9, 10] := 0.000000e+000;
   STAT28[1, 10, 1] := 0.000000e+000;
   STAT28[1, 10, 2] := 0.000000e+000;
   STAT28[1, 10, 3] := 0.000000e+000;
   STAT28[1, 10, 4] := 0.000000e+000;
   STAT28[1, 10, 5] := 0.000000e+000;
   STAT28[1, 10, 6] := 0.000000e+000;
   STAT28[1, 10, 7] := 0.000000e+000;
   STAT28[1, 10, 8] := 0.000000e+000;
   STAT28[1, 10, 9] := 0.000000e+000;
   STAT28[1, 10, 10] := 0.000000e+000;
   STAT28[2, 1, 1] := 0.000000e+000;
   STAT28[2, 1, 2] := 0.000000e+000;
   STAT28[2, 1, 3] := 0.000000e+000;
   STAT28[2, 1, 4] := 0.000000e+000;
   STAT28[2, 1, 5] := 0.000000e+000;
   STAT28[2, 1, 6] := 0.000000e+000;
   STAT28[2, 1, 7] := 0.000000e+000;
   STAT28[2, 1, 8] := 0.000000e+000;
   STAT28[2, 1, 9] := 0.000000e+000;
   STAT28[2, 1, 10] := 0.000000e+000;
   STAT28[2, 2, 1] := 0.000000e+000;
   STAT28[2, 2, 2] := 0.000000e+000;
   STAT28[2, 2, 3] := 0.000000e+000;
   STAT28[2, 2, 4] := 0.000000e+000;
   STAT28[2, 2, 5] := 0.000000e+000;
   STAT28[2, 2, 6] := 0.000000e+000;
   STAT28[2, 2, 7] := 0.000000e+000;
   STAT28[2, 2, 8] := 0.000000e+000;
   STAT28[2, 2, 9] := 0.000000e+000;
   STAT28[2, 2, 10] := 0.000000e+000;
   STAT28[2, 3, 1] := 0.000000e+000;
   STAT28[2, 3, 2] := 0.000000e+000;
   STAT28[2, 3, 3] := 0.000000e+000;
   STAT28[2, 3, 4] := 0.000000e+000;
   STAT28[2, 3, 5] := 0.000000e+000;
   STAT28[2, 3, 6] := 0.000000e+000;
   STAT28[2, 3, 7] := 0.000000e+000;
   STAT28[2, 3, 8] := 0.000000e+000;
   STAT28[2, 3, 9] := 0.000000e+000;
   STAT28[2, 3, 10] := 0.000000e+000;
   STAT28[2, 4, 1] := 0.000000e+000;
   STAT28[2, 4, 2] := 0.000000e+000;
   STAT28[2, 4, 3] := 0.000000e+000;
   STAT28[2, 4, 4] := 0.000000e+000;
   STAT28[2, 4, 5] := 0.000000e+000;
   STAT28[2, 4, 6] := 0.000000e+000;
   STAT28[2, 4, 7] := 0.000000e+000;
   STAT28[2, 4, 8] := 0.000000e+000;
   STAT28[2, 4, 9] := 0.000000e+000;
   STAT28[2, 4, 10] := 0.000000e+000;
   STAT28[2, 5, 1] := 0.000000e+000;
   STAT28[2, 5, 2] := 0.000000e+000;
   STAT28[2, 5, 3] := 0.000000e+000;
   STAT28[2, 5, 4] := 0.000000e+000;
   STAT28[2, 5, 5] := 0.000000e+000;
   STAT28[2, 5, 6] := 0.000000e+000;
   STAT28[2, 5, 7] := 0.000000e+000;
   STAT28[2, 5, 8] := 0.000000e+000;
   STAT28[2, 5, 9] := 0.000000e+000;
   STAT28[2, 5, 10] := 0.000000e+000;
   STAT28[2, 6, 1] := 0.000000e+000;
   STAT28[2, 6, 2] := 0.000000e+000;
   STAT28[2, 6, 3] := 0.000000e+000;
   STAT28[2, 6, 4] := 0.000000e+000;
   STAT28[2, 6, 5] := 0.000000e+000;
   STAT28[2, 6, 6] := 0.000000e+000;
   STAT28[2, 6, 7] := 0.000000e+000;
   STAT28[2, 6, 8] := 0.000000e+000;
   STAT28[2, 6, 9] := 0.000000e+000;
   STAT28[2, 6, 10] := 0.000000e+000;
   STAT28[2, 7, 1] := 0.000000e+000;
   STAT28[2, 7, 2] := 0.000000e+000;
   STAT28[2, 7, 3] := 0.000000e+000;
   STAT28[2, 7, 4] := 0.000000e+000;
   STAT28[2, 7, 5] := 0.000000e+000;
   STAT28[2, 7, 6] := 0.000000e+000;
   STAT28[2, 7, 7] := 0.000000e+000;
   STAT28[2, 7, 8] := 0.000000e+000;
   STAT28[2, 7, 9] := 0.000000e+000;
   STAT28[2, 7, 10] := 0.000000e+000;
   STAT28[2, 8, 1] := 0.000000e+000;
   STAT28[2, 8, 2] := 0.000000e+000;
   STAT28[2, 8, 3] := 0.000000e+000;
   STAT28[2, 8, 4] := 0.000000e+000;
   STAT28[2, 8, 5] := 0.000000e+000;
   STAT28[2, 8, 6] := 0.000000e+000;
   STAT28[2, 8, 7] := 0.000000e+000;
   STAT28[2, 8, 8] := 0.000000e+000;
   STAT28[2, 8, 9] := 0.000000e+000;
   STAT28[2, 8, 10] := 0.000000e+000;
   STAT28[2, 9, 1] := 0.000000e+000;
   STAT28[2, 9, 2] := 0.000000e+000;
   STAT28[2, 9, 3] := 0.000000e+000;
   STAT28[2, 9, 4] := 0.000000e+000;
   STAT28[2, 9, 5] := 0.000000e+000;
   STAT28[2, 9, 6] := 0.000000e+000;
   STAT28[2, 9, 7] := 0.000000e+000;
   STAT28[2, 9, 8] := 0.000000e+000;
   STAT28[2, 9, 9] := 0.000000e+000;
   STAT28[2, 9, 10] := 0.000000e+000;
   STAT28[2, 10, 1] := 0.000000e+000;
   STAT28[2, 10, 2] := 0.000000e+000;
   STAT28[2, 10, 3] := 0.000000e+000;
   STAT28[2, 10, 4] := 0.000000e+000;
   STAT28[2, 10, 5] := 0.000000e+000;
   STAT28[2, 10, 6] := 0.000000e+000;
   STAT28[2, 10, 7] := 0.000000e+000;
   STAT28[2, 10, 8] := 0.000000e+000;
   STAT28[2, 10, 9] := 0.000000e+000;
   STAT28[2, 10, 10] := 0.000000e+000;
   STAT28[3, 1, 1] := 0.000000e+000;
   STAT28[3, 1, 2] := 0.000000e+000;
   STAT28[3, 1, 3] := 0.000000e+000;
   STAT28[3, 1, 4] := 0.000000e+000;
   STAT28[3, 1, 5] := 0.000000e+000;
   STAT28[3, 1, 6] := 0.000000e+000;
   STAT28[3, 1, 7] := 0.000000e+000;
   STAT28[3, 1, 8] := 0.000000e+000;
   STAT28[3, 1, 9] := 0.000000e+000;
   STAT28[3, 1, 10] := 0.000000e+000;
   STAT28[3, 2, 1] := 0.000000e+000;
   STAT28[3, 2, 2] := 0.000000e+000;
   STAT28[3, 2, 3] := 0.000000e+000;
   STAT28[3, 2, 4] := 0.000000e+000;
   STAT28[3, 2, 5] := 0.000000e+000;
   STAT28[3, 2, 6] := 0.000000e+000;
   STAT28[3, 2, 7] := 0.000000e+000;
   STAT28[3, 2, 8] := 0.000000e+000;
   STAT28[3, 2, 9] := 0.000000e+000;
   STAT28[3, 2, 10] := 0.000000e+000;
   STAT28[3, 3, 1] := 0.000000e+000;
   STAT28[3, 3, 2] := 0.000000e+000;
   STAT28[3, 3, 3] := 0.000000e+000;
   STAT28[3, 3, 4] := 0.000000e+000;
   STAT28[3, 3, 5] := 0.000000e+000;
   STAT28[3, 3, 6] := 0.000000e+000;
   STAT28[3, 3, 7] := 0.000000e+000;
   STAT28[3, 3, 8] := 0.000000e+000;
   STAT28[3, 3, 9] := 0.000000e+000;
   STAT28[3, 3, 10] := 0.000000e+000;
   STAT28[3, 4, 1] := 0.000000e+000;
   STAT28[3, 4, 2] := 0.000000e+000;
   STAT28[3, 4, 3] := 0.000000e+000;
   STAT28[3, 4, 4] := 0.000000e+000;
   STAT28[3, 4, 5] := 0.000000e+000;
   STAT28[3, 4, 6] := 0.000000e+000;
   STAT28[3, 4, 7] := 0.000000e+000;
   STAT28[3, 4, 8] := 0.000000e+000;
   STAT28[3, 4, 9] := 0.000000e+000;
   STAT28[3, 4, 10] := 0.000000e+000;
   STAT28[3, 5, 1] := 0.000000e+000;
   STAT28[3, 5, 2] := 0.000000e+000;
   STAT28[3, 5, 3] := 0.000000e+000;
   STAT28[3, 5, 4] := 0.000000e+000;
   STAT28[3, 5, 5] := 0.000000e+000;
   STAT28[3, 5, 6] := 0.000000e+000;
   STAT28[3, 5, 7] := 0.000000e+000;
   STAT28[3, 5, 8] := 0.000000e+000;
   STAT28[3, 5, 9] := 0.000000e+000;
   STAT28[3, 5, 10] := 0.000000e+000;
   STAT28[3, 6, 1] := 0.000000e+000;
   STAT28[3, 6, 2] := 0.000000e+000;
   STAT28[3, 6, 3] := 0.000000e+000;
   STAT28[3, 6, 4] := 0.000000e+000;
   STAT28[3, 6, 5] := 0.000000e+000;
   STAT28[3, 6, 6] := 0.000000e+000;
   STAT28[3, 6, 7] := 0.000000e+000;
   STAT28[3, 6, 8] := 0.000000e+000;
   STAT28[3, 6, 9] := 0.000000e+000;
   STAT28[3, 6, 10] := 0.000000e+000;
   STAT28[3, 7, 1] := 0.000000e+000;
   STAT28[3, 7, 2] := 0.000000e+000;
   STAT28[3, 7, 3] := 0.000000e+000;
   STAT28[3, 7, 4] := 0.000000e+000;
   STAT28[3, 7, 5] := 0.000000e+000;
   STAT28[3, 7, 6] := 0.000000e+000;
   STAT28[3, 7, 7] := 0.000000e+000;
   STAT28[3, 7, 8] := 0.000000e+000;
   STAT28[3, 7, 9] := 0.000000e+000;
   STAT28[3, 7, 10] := 0.000000e+000;
   STAT28[3, 8, 1] := 0.000000e+000;
   STAT28[3, 8, 2] := 0.000000e+000;
   STAT28[3, 8, 3] := 0.000000e+000;
   STAT28[3, 8, 4] := 0.000000e+000;
   STAT28[3, 8, 5] := 0.000000e+000;
   STAT28[3, 8, 6] := 0.000000e+000;
   STAT28[3, 8, 7] := 0.000000e+000;
   STAT28[3, 8, 8] := 0.000000e+000;
   STAT28[3, 8, 9] := 0.000000e+000;
   STAT28[3, 8, 10] := 0.000000e+000;
   STAT28[3, 9, 1] := 0.000000e+000;
   STAT28[3, 9, 2] := 0.000000e+000;
   STAT28[3, 9, 3] := 0.000000e+000;
   STAT28[3, 9, 4] := 0.000000e+000;
   STAT28[3, 9, 5] := 0.000000e+000;
   STAT28[3, 9, 6] := 0.000000e+000;
   STAT28[3, 9, 7] := 0.000000e+000;
   STAT28[3, 9, 8] := 0.000000e+000;
   STAT28[3, 9, 9] := 0.000000e+000;
   STAT28[3, 9, 10] := 0.000000e+000;
   STAT28[3, 10, 1] := 0.000000e+000;
   STAT28[3, 10, 2] := 0.000000e+000;
   STAT28[3, 10, 3] := 0.000000e+000;
   STAT28[3, 10, 4] := 0.000000e+000;
   STAT28[3, 10, 5] := 0.000000e+000;
   STAT28[3, 10, 6] := 0.000000e+000;
   STAT28[3, 10, 7] := 0.000000e+000;
   STAT28[3, 10, 8] := 0.000000e+000;
   STAT28[3, 10, 9] := 0.000000e+000;
   STAT28[3, 10, 10] := 0.000000e+000;
   STAT28[4, 1, 1] := 0.000000e+000;
   STAT28[4, 1, 2] := 0.000000e+000;
   STAT28[4, 1, 3] := 0.000000e+000;
   STAT28[4, 1, 4] := 0.000000e+000;
   STAT28[4, 1, 5] := 0.000000e+000;
   STAT28[4, 1, 6] := 0.000000e+000;
   STAT28[4, 1, 7] := 0.000000e+000;
   STAT28[4, 1, 8] := 0.000000e+000;
   STAT28[4, 1, 9] := 0.000000e+000;
   STAT28[4, 1, 10] := 0.000000e+000;
   STAT28[4, 2, 1] := 0.000000e+000;
   STAT28[4, 2, 2] := 0.000000e+000;
   STAT28[4, 2, 3] := 0.000000e+000;
   STAT28[4, 2, 4] := 0.000000e+000;
   STAT28[4, 2, 5] := 0.000000e+000;
   STAT28[4, 2, 6] := 0.000000e+000;
   STAT28[4, 2, 7] := 0.000000e+000;
   STAT28[4, 2, 8] := 0.000000e+000;
   STAT28[4, 2, 9] := 0.000000e+000;
   STAT28[4, 2, 10] := 0.000000e+000;
   STAT28[4, 3, 1] := 0.000000e+000;
   STAT28[4, 3, 2] := 0.000000e+000;
   STAT28[4, 3, 3] := 0.000000e+000;
   STAT28[4, 3, 4] := 0.000000e+000;
   STAT28[4, 3, 5] := 0.000000e+000;
   STAT28[4, 3, 6] := 0.000000e+000;
   STAT28[4, 3, 7] := 0.000000e+000;
   STAT28[4, 3, 8] := 0.000000e+000;
   STAT28[4, 3, 9] := 0.000000e+000;
   STAT28[4, 3, 10] := 0.000000e+000;
   STAT28[4, 4, 1] := 0.000000e+000;
   STAT28[4, 4, 2] := 0.000000e+000;
   STAT28[4, 4, 3] := 0.000000e+000;
   STAT28[4, 4, 4] := 0.000000e+000;
   STAT28[4, 4, 5] := 0.000000e+000;
   STAT28[4, 4, 6] := 0.000000e+000;
   STAT28[4, 4, 7] := 0.000000e+000;
   STAT28[4, 4, 8] := 0.000000e+000;
   STAT28[4, 4, 9] := 0.000000e+000;
   STAT28[4, 4, 10] := 0.000000e+000;
   STAT28[4, 5, 1] := 0.000000e+000;
   STAT28[4, 5, 2] := 0.000000e+000;
   STAT28[4, 5, 3] := 0.000000e+000;
   STAT28[4, 5, 4] := 0.000000e+000;
   STAT28[4, 5, 5] := 0.000000e+000;
   STAT28[4, 5, 6] := 0.000000e+000;
   STAT28[4, 5, 7] := 0.000000e+000;
   STAT28[4, 5, 8] := 0.000000e+000;
   STAT28[4, 5, 9] := 0.000000e+000;
   STAT28[4, 5, 10] := 0.000000e+000;
   STAT28[4, 6, 1] := 0.000000e+000;
   STAT28[4, 6, 2] := 0.000000e+000;
   STAT28[4, 6, 3] := 0.000000e+000;
   STAT28[4, 6, 4] := 0.000000e+000;
   STAT28[4, 6, 5] := 0.000000e+000;
   STAT28[4, 6, 6] := 0.000000e+000;
   STAT28[4, 6, 7] := 0.000000e+000;
   STAT28[4, 6, 8] := 0.000000e+000;
   STAT28[4, 6, 9] := 0.000000e+000;
   STAT28[4, 6, 10] := 0.000000e+000;
   STAT28[4, 7, 1] := 0.000000e+000;
   STAT28[4, 7, 2] := 0.000000e+000;
   STAT28[4, 7, 3] := 0.000000e+000;
   STAT28[4, 7, 4] := 0.000000e+000;
   STAT28[4, 7, 5] := 0.000000e+000;
   STAT28[4, 7, 6] := 0.000000e+000;
   STAT28[4, 7, 7] := 0.000000e+000;
   STAT28[4, 7, 8] := 0.000000e+000;
   STAT28[4, 7, 9] := 0.000000e+000;
   STAT28[4, 7, 10] := 0.000000e+000;
   STAT28[4, 8, 1] := 0.000000e+000;
   STAT28[4, 8, 2] := 0.000000e+000;
   STAT28[4, 8, 3] := 0.000000e+000;
   STAT28[4, 8, 4] := 0.000000e+000;
   STAT28[4, 8, 5] := 0.000000e+000;
   STAT28[4, 8, 6] := 0.000000e+000;
   STAT28[4, 8, 7] := 0.000000e+000;
   STAT28[4, 8, 8] := 0.000000e+000;
   STAT28[4, 8, 9] := 0.000000e+000;
   STAT28[4, 8, 10] := 0.000000e+000;
   STAT28[4, 9, 1] := 0.000000e+000;
   STAT28[4, 9, 2] := 0.000000e+000;
   STAT28[4, 9, 3] := 0.000000e+000;
   STAT28[4, 9, 4] := 0.000000e+000;
   STAT28[4, 9, 5] := 0.000000e+000;
   STAT28[4, 9, 6] := 0.000000e+000;
   STAT28[4, 9, 7] := 0.000000e+000;
   STAT28[4, 9, 8] := 0.000000e+000;
   STAT28[4, 9, 9] := 0.000000e+000;
   STAT28[4, 9, 10] := 0.000000e+000;
   STAT28[4, 10, 1] := 0.000000e+000;
   STAT28[4, 10, 2] := 0.000000e+000;
   STAT28[4, 10, 3] := 0.000000e+000;
   STAT28[4, 10, 4] := 0.000000e+000;
   STAT28[4, 10, 5] := 0.000000e+000;
   STAT28[4, 10, 6] := 0.000000e+000;
   STAT28[4, 10, 7] := 0.000000e+000;
   STAT28[4, 10, 8] := 0.000000e+000;
   STAT28[4, 10, 9] := 0.000000e+000;
   STAT28[4, 10, 10] := 0.000000e+000;
   STAT28[5, 1, 1] := 0.000000e+000;
   STAT28[5, 1, 2] := 0.000000e+000;
   STAT28[5, 1, 3] := 0.000000e+000;
   STAT28[5, 1, 4] := 0.000000e+000;
   STAT28[5, 1, 5] := 0.000000e+000;
   STAT28[5, 1, 6] := 0.000000e+000;
   STAT28[5, 1, 7] := 0.000000e+000;
   STAT28[5, 1, 8] := 0.000000e+000;
   STAT28[5, 1, 9] := 0.000000e+000;
   STAT28[5, 1, 10] := 0.000000e+000;
   STAT28[5, 2, 1] := 0.000000e+000;
   STAT28[5, 2, 2] := 0.000000e+000;
   STAT28[5, 2, 3] := 0.000000e+000;
   STAT28[5, 2, 4] := 0.000000e+000;
   STAT28[5, 2, 5] := 0.000000e+000;
   STAT28[5, 2, 6] := 0.000000e+000;
   STAT28[5, 2, 7] := 0.000000e+000;
   STAT28[5, 2, 8] := 0.000000e+000;
   STAT28[5, 2, 9] := 0.000000e+000;
   STAT28[5, 2, 10] := 0.000000e+000;
   STAT28[5, 3, 1] := 0.000000e+000;
   STAT28[5, 3, 2] := 0.000000e+000;
   STAT28[5, 3, 3] := 0.000000e+000;
   STAT28[5, 3, 4] := 0.000000e+000;
   STAT28[5, 3, 5] := 0.000000e+000;
   STAT28[5, 3, 6] := 0.000000e+000;
   STAT28[5, 3, 7] := 0.000000e+000;
   STAT28[5, 3, 8] := 0.000000e+000;
   STAT28[5, 3, 9] := 0.000000e+000;
   STAT28[5, 3, 10] := 0.000000e+000;
   STAT28[5, 4, 1] := 0.000000e+000;
   STAT28[5, 4, 2] := 0.000000e+000;
   STAT28[5, 4, 3] := 0.000000e+000;
   STAT28[5, 4, 4] := 0.000000e+000;
   STAT28[5, 4, 5] := 0.000000e+000;
   STAT28[5, 4, 6] := 0.000000e+000;
   STAT28[5, 4, 7] := 0.000000e+000;
   STAT28[5, 4, 8] := 0.000000e+000;
   STAT28[5, 4, 9] := 0.000000e+000;
   STAT28[5, 4, 10] := 0.000000e+000;
   STAT28[5, 5, 1] := 0.000000e+000;
   STAT28[5, 5, 2] := 0.000000e+000;
   STAT28[5, 5, 3] := 0.000000e+000;
   STAT28[5, 5, 4] := 0.000000e+000;
   STAT28[5, 5, 5] := 0.000000e+000;
   STAT28[5, 5, 6] := 0.000000e+000;
   STAT28[5, 5, 7] := 0.000000e+000;
   STAT28[5, 5, 8] := 0.000000e+000;
   STAT28[5, 5, 9] := 0.000000e+000;
   STAT28[5, 5, 10] := 0.000000e+000;
   STAT28[5, 6, 1] := 0.000000e+000;
   STAT28[5, 6, 2] := 0.000000e+000;
   STAT28[5, 6, 3] := 0.000000e+000;
   STAT28[5, 6, 4] := 0.000000e+000;
   STAT28[5, 6, 5] := 0.000000e+000;
   STAT28[5, 6, 6] := 0.000000e+000;
   STAT28[5, 6, 7] := 0.000000e+000;
   STAT28[5, 6, 8] := 0.000000e+000;
   STAT28[5, 6, 9] := 0.000000e+000;
   STAT28[5, 6, 10] := 0.000000e+000;
   STAT28[5, 7, 1] := 0.000000e+000;
   STAT28[5, 7, 2] := 0.000000e+000;
   STAT28[5, 7, 3] := 0.000000e+000;
   STAT28[5, 7, 4] := 0.000000e+000;
   STAT28[5, 7, 5] := 0.000000e+000;
   STAT28[5, 7, 6] := 0.000000e+000;
   STAT28[5, 7, 7] := 0.000000e+000;
   STAT28[5, 7, 8] := 0.000000e+000;
   STAT28[5, 7, 9] := 0.000000e+000;
   STAT28[5, 7, 10] := 0.000000e+000;
   STAT28[5, 8, 1] := 0.000000e+000;
   STAT28[5, 8, 2] := 0.000000e+000;
   STAT28[5, 8, 3] := 0.000000e+000;
   STAT28[5, 8, 4] := 0.000000e+000;
   STAT28[5, 8, 5] := 0.000000e+000;
   STAT28[5, 8, 6] := 0.000000e+000;
   STAT28[5, 8, 7] := 0.000000e+000;
   STAT28[5, 8, 8] := 0.000000e+000;
   STAT28[5, 8, 9] := 0.000000e+000;
   STAT28[5, 8, 10] := 0.000000e+000;
   STAT28[5, 9, 1] := 0.000000e+000;
   STAT28[5, 9, 2] := 0.000000e+000;
   STAT28[5, 9, 3] := 0.000000e+000;
   STAT28[5, 9, 4] := 0.000000e+000;
   STAT28[5, 9, 5] := 0.000000e+000;
   STAT28[5, 9, 6] := 0.000000e+000;
   STAT28[5, 9, 7] := 0.000000e+000;
   STAT28[5, 9, 8] := 0.000000e+000;
   STAT28[5, 9, 9] := 0.000000e+000;
   STAT28[5, 9, 10] := 0.000000e+000;
   STAT28[5, 10, 1] := 0.000000e+000;
   STAT28[5, 10, 2] := 0.000000e+000;
   STAT28[5, 10, 3] := 0.000000e+000;
   STAT28[5, 10, 4] := 0.000000e+000;
   STAT28[5, 10, 5] := 0.000000e+000;
   STAT28[5, 10, 6] := 0.000000e+000;
   STAT28[5, 10, 7] := 0.000000e+000;
   STAT28[5, 10, 8] := 0.000000e+000;
   STAT28[5, 10, 9] := 0.000000e+000;
   STAT28[5, 10, 10] := 0.000000e+000;
   STAT28[6, 1, 1] := 0.000000e+000;
   STAT28[6, 1, 2] := 0.000000e+000;
   STAT28[6, 1, 3] := 0.000000e+000;
   STAT28[6, 1, 4] := 0.000000e+000;
   STAT28[6, 1, 5] := 0.000000e+000;
   STAT28[6, 1, 6] := 0.000000e+000;
   STAT28[6, 1, 7] := 0.000000e+000;
   STAT28[6, 1, 8] := 0.000000e+000;
   STAT28[6, 1, 9] := 0.000000e+000;
   STAT28[6, 1, 10] := 0.000000e+000;
   STAT28[6, 2, 1] := 0.000000e+000;
   STAT28[6, 2, 2] := 0.000000e+000;
   STAT28[6, 2, 3] := 0.000000e+000;
   STAT28[6, 2, 4] := 0.000000e+000;
   STAT28[6, 2, 5] := 0.000000e+000;
   STAT28[6, 2, 6] := 0.000000e+000;
   STAT28[6, 2, 7] := 0.000000e+000;
   STAT28[6, 2, 8] := 0.000000e+000;
   STAT28[6, 2, 9] := 0.000000e+000;
   STAT28[6, 2, 10] := 0.000000e+000;
   STAT28[6, 3, 1] := 0.000000e+000;
   STAT28[6, 3, 2] := 0.000000e+000;
   STAT28[6, 3, 3] := 0.000000e+000;
   STAT28[6, 3, 4] := 0.000000e+000;
   STAT28[6, 3, 5] := 0.000000e+000;
   STAT28[6, 3, 6] := 0.000000e+000;
   STAT28[6, 3, 7] := 0.000000e+000;
   STAT28[6, 3, 8] := 0.000000e+000;
   STAT28[6, 3, 9] := 0.000000e+000;
   STAT28[6, 3, 10] := 0.000000e+000;
   STAT28[6, 4, 1] := 0.000000e+000;
   STAT28[6, 4, 2] := 0.000000e+000;
   STAT28[6, 4, 3] := 0.000000e+000;
   STAT28[6, 4, 4] := 0.000000e+000;
   STAT28[6, 4, 5] := 0.000000e+000;
   STAT28[6, 4, 6] := 0.000000e+000;
   STAT28[6, 4, 7] := 0.000000e+000;
   STAT28[6, 4, 8] := 0.000000e+000;
   STAT28[6, 4, 9] := 0.000000e+000;
   STAT28[6, 4, 10] := 0.000000e+000;
   STAT28[6, 5, 1] := 0.000000e+000;
   STAT28[6, 5, 2] := 0.000000e+000;
   STAT28[6, 5, 3] := 0.000000e+000;
   STAT28[6, 5, 4] := 0.000000e+000;
   STAT28[6, 5, 5] := 0.000000e+000;
   STAT28[6, 5, 6] := 0.000000e+000;
   STAT28[6, 5, 7] := 0.000000e+000;
   STAT28[6, 5, 8] := 0.000000e+000;
   STAT28[6, 5, 9] := 0.000000e+000;
   STAT28[6, 5, 10] := 0.000000e+000;
   STAT28[6, 6, 1] := 0.000000e+000;
   STAT28[6, 6, 2] := 0.000000e+000;
   STAT28[6, 6, 3] := 0.000000e+000;
   STAT28[6, 6, 4] := 0.000000e+000;
   STAT28[6, 6, 5] := 0.000000e+000;
   STAT28[6, 6, 6] := 0.000000e+000;
   STAT28[6, 6, 7] := 0.000000e+000;
   STAT28[6, 6, 8] := 0.000000e+000;
   STAT28[6, 6, 9] := 0.000000e+000;
   STAT28[6, 6, 10] := 0.000000e+000;
   STAT28[6, 7, 1] := 0.000000e+000;
   STAT28[6, 7, 2] := 0.000000e+000;
   STAT28[6, 7, 3] := 0.000000e+000;
   STAT28[6, 7, 4] := 0.000000e+000;
   STAT28[6, 7, 5] := 0.000000e+000;
   STAT28[6, 7, 6] := 0.000000e+000;
   STAT28[6, 7, 7] := 0.000000e+000;
   STAT28[6, 7, 8] := 0.000000e+000;
   STAT28[6, 7, 9] := 0.000000e+000;
   STAT28[6, 7, 10] := 0.000000e+000;
   STAT28[6, 8, 1] := 0.000000e+000;
   STAT28[6, 8, 2] := 0.000000e+000;
   STAT28[6, 8, 3] := 0.000000e+000;
   STAT28[6, 8, 4] := 0.000000e+000;
   STAT28[6, 8, 5] := 0.000000e+000;
   STAT28[6, 8, 6] := 0.000000e+000;
   STAT28[6, 8, 7] := 0.000000e+000;
   STAT28[6, 8, 8] := 0.000000e+000;
   STAT28[6, 8, 9] := 0.000000e+000;
   STAT28[6, 8, 10] := 0.000000e+000;
   STAT28[6, 9, 1] := 0.000000e+000;
   STAT28[6, 9, 2] := 0.000000e+000;
   STAT28[6, 9, 3] := 0.000000e+000;
   STAT28[6, 9, 4] := 0.000000e+000;
   STAT28[6, 9, 5] := 0.000000e+000;
   STAT28[6, 9, 6] := 0.000000e+000;
   STAT28[6, 9, 7] := 0.000000e+000;
   STAT28[6, 9, 8] := 0.000000e+000;
   STAT28[6, 9, 9] := 0.000000e+000;
   STAT28[6, 9, 10] := 0.000000e+000;
   STAT28[6, 10, 1] := 0.000000e+000;
   STAT28[6, 10, 2] := 0.000000e+000;
   STAT28[6, 10, 3] := 0.000000e+000;
   STAT28[6, 10, 4] := 0.000000e+000;
   STAT28[6, 10, 5] := 0.000000e+000;
   STAT28[6, 10, 6] := 0.000000e+000;
   STAT28[6, 10, 7] := 0.000000e+000;
   STAT28[6, 10, 8] := 0.000000e+000;
   STAT28[6, 10, 9] := 0.000000e+000;
   STAT28[6, 10, 10] := 0.000000e+000;
   STAT28[7, 1, 1] := 0.000000e+000;
   STAT28[7, 1, 2] := 0.000000e+000;
   STAT28[7, 1, 3] := 0.000000e+000;
   STAT28[7, 1, 4] := 0.000000e+000;
   STAT28[7, 1, 5] := 0.000000e+000;
   STAT28[7, 1, 6] := 0.000000e+000;
   STAT28[7, 1, 7] := 0.000000e+000;
   STAT28[7, 1, 8] := 0.000000e+000;
   STAT28[7, 1, 9] := 0.000000e+000;
   STAT28[7, 1, 10] := 0.000000e+000;
   STAT28[7, 2, 1] := 0.000000e+000;
   STAT28[7, 2, 2] := 0.000000e+000;
   STAT28[7, 2, 3] := 0.000000e+000;
   STAT28[7, 2, 4] := 0.000000e+000;
   STAT28[7, 2, 5] := 0.000000e+000;
   STAT28[7, 2, 6] := 0.000000e+000;
   STAT28[7, 2, 7] := 0.000000e+000;
   STAT28[7, 2, 8] := 0.000000e+000;
   STAT28[7, 2, 9] := 0.000000e+000;
   STAT28[7, 2, 10] := 0.000000e+000;
   STAT28[7, 3, 1] := 0.000000e+000;
   STAT28[7, 3, 2] := 0.000000e+000;
   STAT28[7, 3, 3] := 0.000000e+000;
   STAT28[7, 3, 4] := 0.000000e+000;
   STAT28[7, 3, 5] := 0.000000e+000;
   STAT28[7, 3, 6] := 0.000000e+000;
   STAT28[7, 3, 7] := 0.000000e+000;
   STAT28[7, 3, 8] := 0.000000e+000;
   STAT28[7, 3, 9] := 0.000000e+000;
   STAT28[7, 3, 10] := 0.000000e+000;
   STAT28[7, 4, 1] := 0.000000e+000;
   STAT28[7, 4, 2] := 0.000000e+000;
   STAT28[7, 4, 3] := 0.000000e+000;
   STAT28[7, 4, 4] := 0.000000e+000;
   STAT28[7, 4, 5] := 0.000000e+000;
   STAT28[7, 4, 6] := 0.000000e+000;
   STAT28[7, 4, 7] := 0.000000e+000;
   STAT28[7, 4, 8] := 0.000000e+000;
   STAT28[7, 4, 9] := 0.000000e+000;
   STAT28[7, 4, 10] := 0.000000e+000;
   STAT28[7, 5, 1] := 0.000000e+000;
   STAT28[7, 5, 2] := 0.000000e+000;
   STAT28[7, 5, 3] := 0.000000e+000;
   STAT28[7, 5, 4] := 0.000000e+000;
   STAT28[7, 5, 5] := 0.000000e+000;
   STAT28[7, 5, 6] := 0.000000e+000;
   STAT28[7, 5, 7] := 0.000000e+000;
   STAT28[7, 5, 8] := 0.000000e+000;
   STAT28[7, 5, 9] := 0.000000e+000;
   STAT28[7, 5, 10] := 0.000000e+000;
   STAT28[7, 6, 1] := 0.000000e+000;
   STAT28[7, 6, 2] := 0.000000e+000;
   STAT28[7, 6, 3] := 0.000000e+000;
   STAT28[7, 6, 4] := 0.000000e+000;
   STAT28[7, 6, 5] := 0.000000e+000;
   STAT28[7, 6, 6] := 0.000000e+000;
   STAT28[7, 6, 7] := 0.000000e+000;
   STAT28[7, 6, 8] := 0.000000e+000;
   STAT28[7, 6, 9] := 0.000000e+000;
   STAT28[7, 6, 10] := 0.000000e+000;
   STAT28[7, 7, 1] := 0.000000e+000;
   STAT28[7, 7, 2] := 0.000000e+000;
   STAT28[7, 7, 3] := 0.000000e+000;
   STAT28[7, 7, 4] := 0.000000e+000;
   STAT28[7, 7, 5] := 0.000000e+000;
   STAT28[7, 7, 6] := 0.000000e+000;
   STAT28[7, 7, 7] := 0.000000e+000;
   STAT28[7, 7, 8] := 0.000000e+000;
   STAT28[7, 7, 9] := 0.000000e+000;
   STAT28[7, 7, 10] := 0.000000e+000;
   STAT28[7, 8, 1] := 0.000000e+000;
   STAT28[7, 8, 2] := 0.000000e+000;
   STAT28[7, 8, 3] := 0.000000e+000;
   STAT28[7, 8, 4] := 0.000000e+000;
   STAT28[7, 8, 5] := 0.000000e+000;
   STAT28[7, 8, 6] := 0.000000e+000;
   STAT28[7, 8, 7] := 0.000000e+000;
   STAT28[7, 8, 8] := 0.000000e+000;
   STAT28[7, 8, 9] := 0.000000e+000;
   STAT28[7, 8, 10] := 0.000000e+000;
   STAT28[7, 9, 1] := 0.000000e+000;
   STAT28[7, 9, 2] := 0.000000e+000;
   STAT28[7, 9, 3] := 0.000000e+000;
   STAT28[7, 9, 4] := 0.000000e+000;
   STAT28[7, 9, 5] := 0.000000e+000;
   STAT28[7, 9, 6] := 0.000000e+000;
   STAT28[7, 9, 7] := 0.000000e+000;
   STAT28[7, 9, 8] := 0.000000e+000;
   STAT28[7, 9, 9] := 0.000000e+000;
   STAT28[7, 9, 10] := 0.000000e+000;
   STAT28[7, 10, 1] := 0.000000e+000;
   STAT28[7, 10, 2] := 0.000000e+000;
   STAT28[7, 10, 3] := 0.000000e+000;
   STAT28[7, 10, 4] := 0.000000e+000;
   STAT28[7, 10, 5] := 0.000000e+000;
   STAT28[7, 10, 6] := 0.000000e+000;
   STAT28[7, 10, 7] := 0.000000e+000;
   STAT28[7, 10, 8] := 0.000000e+000;
   STAT28[7, 10, 9] := 0.000000e+000;
   STAT28[7, 10, 10] := 0.000000e+000;
   STAT28[8, 1, 1] := 0.000000e+000;
   STAT28[8, 1, 2] := 0.000000e+000;
   STAT28[8, 1, 3] := 0.000000e+000;
   STAT28[8, 1, 4] := 0.000000e+000;
   STAT28[8, 1, 5] := 0.000000e+000;
   STAT28[8, 1, 6] := 0.000000e+000;
   STAT28[8, 1, 7] := 0.000000e+000;
   STAT28[8, 1, 8] := 0.000000e+000;
   STAT28[8, 1, 9] := 0.000000e+000;
   STAT28[8, 1, 10] := 0.000000e+000;
   STAT28[8, 2, 1] := 0.000000e+000;
   STAT28[8, 2, 2] := 0.000000e+000;
   STAT28[8, 2, 3] := 0.000000e+000;
   STAT28[8, 2, 4] := 0.000000e+000;
   STAT28[8, 2, 5] := 0.000000e+000;
   STAT28[8, 2, 6] := 0.000000e+000;
   STAT28[8, 2, 7] := 0.000000e+000;
   STAT28[8, 2, 8] := 0.000000e+000;
   STAT28[8, 2, 9] := 0.000000e+000;
   STAT28[8, 2, 10] := 0.000000e+000;
   STAT28[8, 3, 1] := 0.000000e+000;
   STAT28[8, 3, 2] := 0.000000e+000;
   STAT28[8, 3, 3] := 0.000000e+000;
   STAT28[8, 3, 4] := 0.000000e+000;
   STAT28[8, 3, 5] := 0.000000e+000;
   STAT28[8, 3, 6] := 0.000000e+000;
   STAT28[8, 3, 7] := 0.000000e+000;
   STAT28[8, 3, 8] := 0.000000e+000;
   STAT28[8, 3, 9] := 0.000000e+000;
   STAT28[8, 3, 10] := 0.000000e+000;
   STAT28[8, 4, 1] := 0.000000e+000;
   STAT28[8, 4, 2] := 0.000000e+000;
   STAT28[8, 4, 3] := 0.000000e+000;
   STAT28[8, 4, 4] := 0.000000e+000;
   STAT28[8, 4, 5] := 0.000000e+000;
   STAT28[8, 4, 6] := 0.000000e+000;
   STAT28[8, 4, 7] := 0.000000e+000;
   STAT28[8, 4, 8] := 0.000000e+000;
   STAT28[8, 4, 9] := 0.000000e+000;
   STAT28[8, 4, 10] := 0.000000e+000;
   STAT28[8, 5, 1] := 0.000000e+000;
   STAT28[8, 5, 2] := 0.000000e+000;
   STAT28[8, 5, 3] := 0.000000e+000;
   STAT28[8, 5, 4] := 0.000000e+000;
   STAT28[8, 5, 5] := 0.000000e+000;
   STAT28[8, 5, 6] := 0.000000e+000;
   STAT28[8, 5, 7] := 0.000000e+000;
   STAT28[8, 5, 8] := 0.000000e+000;
   STAT28[8, 5, 9] := 0.000000e+000;
   STAT28[8, 5, 10] := 0.000000e+000;
   STAT28[8, 6, 1] := 0.000000e+000;
   STAT28[8, 6, 2] := 0.000000e+000;
   STAT28[8, 6, 3] := 0.000000e+000;
   STAT28[8, 6, 4] := 0.000000e+000;
   STAT28[8, 6, 5] := 0.000000e+000;
   STAT28[8, 6, 6] := 0.000000e+000;
   STAT28[8, 6, 7] := 0.000000e+000;
   STAT28[8, 6, 8] := 0.000000e+000;
   STAT28[8, 6, 9] := 0.000000e+000;
   STAT28[8, 6, 10] := 0.000000e+000;
   STAT28[8, 7, 1] := 0.000000e+000;
   STAT28[8, 7, 2] := 0.000000e+000;
   STAT28[8, 7, 3] := 0.000000e+000;
   STAT28[8, 7, 4] := 0.000000e+000;
   STAT28[8, 7, 5] := 0.000000e+000;
   STAT28[8, 7, 6] := 0.000000e+000;
   STAT28[8, 7, 7] := 0.000000e+000;
   STAT28[8, 7, 8] := 0.000000e+000;
   STAT28[8, 7, 9] := 0.000000e+000;
   STAT28[8, 7, 10] := 0.000000e+000;
   STAT28[8, 8, 1] := 0.000000e+000;
   STAT28[8, 8, 2] := 0.000000e+000;
   STAT28[8, 8, 3] := 0.000000e+000;
   STAT28[8, 8, 4] := 0.000000e+000;
   STAT28[8, 8, 5] := 0.000000e+000;
   STAT28[8, 8, 6] := 0.000000e+000;
   STAT28[8, 8, 7] := 0.000000e+000;
   STAT28[8, 8, 8] := 0.000000e+000;
   STAT28[8, 8, 9] := 0.000000e+000;
   STAT28[8, 8, 10] := 0.000000e+000;
   STAT28[8, 9, 1] := 0.000000e+000;
   STAT28[8, 9, 2] := 0.000000e+000;
   STAT28[8, 9, 3] := 0.000000e+000;
   STAT28[8, 9, 4] := 0.000000e+000;
   STAT28[8, 9, 5] := 0.000000e+000;
   STAT28[8, 9, 6] := 0.000000e+000;
   STAT28[8, 9, 7] := 0.000000e+000;
   STAT28[8, 9, 8] := 0.000000e+000;
   STAT28[8, 9, 9] := 0.000000e+000;
   STAT28[8, 9, 10] := 0.000000e+000;
   STAT28[8, 10, 1] := 0.000000e+000;
   STAT28[8, 10, 2] := 0.000000e+000;
   STAT28[8, 10, 3] := 0.000000e+000;
   STAT28[8, 10, 4] := 0.000000e+000;
   STAT28[8, 10, 5] := 0.000000e+000;
   STAT28[8, 10, 6] := 0.000000e+000;
   STAT28[8, 10, 7] := 0.000000e+000;
   STAT28[8, 10, 8] := 0.000000e+000;
   STAT28[8, 10, 9] := 0.000000e+000;
   STAT28[8, 10, 10] := 0.000000e+000;
   STAT28[9, 1, 1] := 0.000000e+000;
   STAT28[9, 1, 2] := 0.000000e+000;
   STAT28[9, 1, 3] := 0.000000e+000;
   STAT28[9, 1, 4] := 0.000000e+000;
   STAT28[9, 1, 5] := 0.000000e+000;
   STAT28[9, 1, 6] := 0.000000e+000;
   STAT28[9, 1, 7] := 0.000000e+000;
   STAT28[9, 1, 8] := 0.000000e+000;
   STAT28[9, 1, 9] := 0.000000e+000;
   STAT28[9, 1, 10] := 0.000000e+000;
   STAT28[9, 2, 1] := 0.000000e+000;
   STAT28[9, 2, 2] := 0.000000e+000;
   STAT28[9, 2, 3] := 0.000000e+000;
   STAT28[9, 2, 4] := 0.000000e+000;
   STAT28[9, 2, 5] := 0.000000e+000;
   STAT28[9, 2, 6] := 0.000000e+000;
   STAT28[9, 2, 7] := 0.000000e+000;
   STAT28[9, 2, 8] := 0.000000e+000;
   STAT28[9, 2, 9] := 0.000000e+000;
   STAT28[9, 2, 10] := 0.000000e+000;
   STAT28[9, 3, 1] := 0.000000e+000;
   STAT28[9, 3, 2] := 0.000000e+000;
   STAT28[9, 3, 3] := 0.000000e+000;
   STAT28[9, 3, 4] := 0.000000e+000;
   STAT28[9, 3, 5] := 0.000000e+000;
   STAT28[9, 3, 6] := 0.000000e+000;
   STAT28[9, 3, 7] := 0.000000e+000;
   STAT28[9, 3, 8] := 0.000000e+000;
   STAT28[9, 3, 9] := 0.000000e+000;
   STAT28[9, 3, 10] := 0.000000e+000;
   STAT28[9, 4, 1] := 0.000000e+000;
   STAT28[9, 4, 2] := 0.000000e+000;
   STAT28[9, 4, 3] := 0.000000e+000;
   STAT28[9, 4, 4] := 0.000000e+000;
   STAT28[9, 4, 5] := 0.000000e+000;
   STAT28[9, 4, 6] := 0.000000e+000;
   STAT28[9, 4, 7] := 0.000000e+000;
   STAT28[9, 4, 8] := 0.000000e+000;
   STAT28[9, 4, 9] := 0.000000e+000;
   STAT28[9, 4, 10] := 0.000000e+000;
   STAT28[9, 5, 1] := 0.000000e+000;
   STAT28[9, 5, 2] := 0.000000e+000;
   STAT28[9, 5, 3] := 0.000000e+000;
   STAT28[9, 5, 4] := 0.000000e+000;
   STAT28[9, 5, 5] := 0.000000e+000;
   STAT28[9, 5, 6] := 0.000000e+000;
   STAT28[9, 5, 7] := 0.000000e+000;
   STAT28[9, 5, 8] := 0.000000e+000;
   STAT28[9, 5, 9] := 0.000000e+000;
   STAT28[9, 5, 10] := 0.000000e+000;
   STAT28[9, 6, 1] := 0.000000e+000;
   STAT28[9, 6, 2] := 0.000000e+000;
   STAT28[9, 6, 3] := 0.000000e+000;
   STAT28[9, 6, 4] := 0.000000e+000;
   STAT28[9, 6, 5] := 0.000000e+000;
   STAT28[9, 6, 6] := 0.000000e+000;
   STAT28[9, 6, 7] := 0.000000e+000;
   STAT28[9, 6, 8] := 0.000000e+000;
   STAT28[9, 6, 9] := 0.000000e+000;
   STAT28[9, 6, 10] := 0.000000e+000;
   STAT28[9, 7, 1] := 0.000000e+000;
   STAT28[9, 7, 2] := 0.000000e+000;
   STAT28[9, 7, 3] := 0.000000e+000;
   STAT28[9, 7, 4] := 0.000000e+000;
   STAT28[9, 7, 5] := 0.000000e+000;
   STAT28[9, 7, 6] := 0.000000e+000;
   STAT28[9, 7, 7] := 0.000000e+000;
   STAT28[9, 7, 8] := 0.000000e+000;
   STAT28[9, 7, 9] := 0.000000e+000;
   STAT28[9, 7, 10] := 0.000000e+000;
   STAT28[9, 8, 1] := 0.000000e+000;
   STAT28[9, 8, 2] := 0.000000e+000;
   STAT28[9, 8, 3] := 0.000000e+000;
   STAT28[9, 8, 4] := 0.000000e+000;
   STAT28[9, 8, 5] := 0.000000e+000;
   STAT28[9, 8, 6] := 0.000000e+000;
   STAT28[9, 8, 7] := 0.000000e+000;
   STAT28[9, 8, 8] := 0.000000e+000;
   STAT28[9, 8, 9] := 0.000000e+000;
   STAT28[9, 8, 10] := 0.000000e+000;
   STAT28[9, 9, 1] := 0.000000e+000;
   STAT28[9, 9, 2] := 0.000000e+000;
   STAT28[9, 9, 3] := 0.000000e+000;
   STAT28[9, 9, 4] := 0.000000e+000;
   STAT28[9, 9, 5] := 0.000000e+000;
   STAT28[9, 9, 6] := 0.000000e+000;
   STAT28[9, 9, 7] := 0.000000e+000;
   STAT28[9, 9, 8] := 0.000000e+000;
   STAT28[9, 9, 9] := 0.000000e+000;
   STAT28[9, 9, 10] := 0.000000e+000;
   STAT28[9, 10, 1] := 0.000000e+000;
   STAT28[9, 10, 2] := 0.000000e+000;
   STAT28[9, 10, 3] := 0.000000e+000;
   STAT28[9, 10, 4] := 0.000000e+000;
   STAT28[9, 10, 5] := 0.000000e+000;
   STAT28[9, 10, 6] := 0.000000e+000;
   STAT28[9, 10, 7] := 0.000000e+000;
   STAT28[9, 10, 8] := 0.000000e+000;
   STAT28[9, 10, 9] := 0.000000e+000;
   STAT28[9, 10, 10] := 0.000000e+000;
   STAT28[10, 1, 1] := 0.000000e+000;
   STAT28[10, 1, 2] := 0.000000e+000;
   STAT28[10, 1, 3] := 0.000000e+000;
   STAT28[10, 1, 4] := 0.000000e+000;
   STAT28[10, 1, 5] := 0.000000e+000;
   STAT28[10, 1, 6] := 0.000000e+000;
   STAT28[10, 1, 7] := 0.000000e+000;
   STAT28[10, 1, 8] := 0.000000e+000;
   STAT28[10, 1, 9] := 0.000000e+000;
   STAT28[10, 1, 10] := 0.000000e+000;
   STAT28[10, 2, 1] := 0.000000e+000;
   STAT28[10, 2, 2] := 0.000000e+000;
   STAT28[10, 2, 3] := 0.000000e+000;
   STAT28[10, 2, 4] := 0.000000e+000;
   STAT28[10, 2, 5] := 0.000000e+000;
   STAT28[10, 2, 6] := 0.000000e+000;
   STAT28[10, 2, 7] := 0.000000e+000;
   STAT28[10, 2, 8] := 0.000000e+000;
   STAT28[10, 2, 9] := 0.000000e+000;
   STAT28[10, 2, 10] := 0.000000e+000;
   STAT28[10, 3, 1] := 0.000000e+000;
   STAT28[10, 3, 2] := 0.000000e+000;
   STAT28[10, 3, 3] := 0.000000e+000;
   STAT28[10, 3, 4] := 0.000000e+000;
   STAT28[10, 3, 5] := 0.000000e+000;
   STAT28[10, 3, 6] := 0.000000e+000;
   STAT28[10, 3, 7] := 0.000000e+000;
   STAT28[10, 3, 8] := 0.000000e+000;
   STAT28[10, 3, 9] := 0.000000e+000;
   STAT28[10, 3, 10] := 0.000000e+000;
   STAT28[10, 4, 1] := 0.000000e+000;
   STAT28[10, 4, 2] := 0.000000e+000;
   STAT28[10, 4, 3] := 0.000000e+000;
   STAT28[10, 4, 4] := 0.000000e+000;
   STAT28[10, 4, 5] := 0.000000e+000;
   STAT28[10, 4, 6] := 0.000000e+000;
   STAT28[10, 4, 7] := 0.000000e+000;
   STAT28[10, 4, 8] := 0.000000e+000;
   STAT28[10, 4, 9] := 0.000000e+000;
   STAT28[10, 4, 10] := 0.000000e+000;
   STAT28[10, 5, 1] := 0.000000e+000;
   STAT28[10, 5, 2] := 0.000000e+000;
   STAT28[10, 5, 3] := 0.000000e+000;
   STAT28[10, 5, 4] := 0.000000e+000;
   STAT28[10, 5, 5] := 0.000000e+000;
   STAT28[10, 5, 6] := 0.000000e+000;
   STAT28[10, 5, 7] := 0.000000e+000;
   STAT28[10, 5, 8] := 0.000000e+000;
   STAT28[10, 5, 9] := 0.000000e+000;
   STAT28[10, 5, 10] := 0.000000e+000;
   STAT28[10, 6, 1] := 0.000000e+000;
   STAT28[10, 6, 2] := 0.000000e+000;
   STAT28[10, 6, 3] := 0.000000e+000;
   STAT28[10, 6, 4] := 0.000000e+000;
   STAT28[10, 6, 5] := 0.000000e+000;
   STAT28[10, 6, 6] := 0.000000e+000;
   STAT28[10, 6, 7] := 0.000000e+000;
   STAT28[10, 6, 8] := 0.000000e+000;
   STAT28[10, 6, 9] := 0.000000e+000;
   STAT28[10, 6, 10] := 0.000000e+000;
   STAT28[10, 7, 1] := 0.000000e+000;
   STAT28[10, 7, 2] := 0.000000e+000;
   STAT28[10, 7, 3] := 0.000000e+000;
   STAT28[10, 7, 4] := 0.000000e+000;
   STAT28[10, 7, 5] := 0.000000e+000;
   STAT28[10, 7, 6] := 0.000000e+000;
   STAT28[10, 7, 7] := 0.000000e+000;
   STAT28[10, 7, 8] := 0.000000e+000;
   STAT28[10, 7, 9] := 0.000000e+000;
   STAT28[10, 7, 10] := 0.000000e+000;
   STAT28[10, 8, 1] := 0.000000e+000;
   STAT28[10, 8, 2] := 0.000000e+000;
   STAT28[10, 8, 3] := 0.000000e+000;
   STAT28[10, 8, 4] := 0.000000e+000;
   STAT28[10, 8, 5] := 0.000000e+000;
   STAT28[10, 8, 6] := 0.000000e+000;
   STAT28[10, 8, 7] := 0.000000e+000;
   STAT28[10, 8, 8] := 0.000000e+000;
   STAT28[10, 8, 9] := 0.000000e+000;
   STAT28[10, 8, 10] := 0.000000e+000;
   STAT28[10, 9, 1] := 0.000000e+000;
   STAT28[10, 9, 2] := 0.000000e+000;
   STAT28[10, 9, 3] := 0.000000e+000;
   STAT28[10, 9, 4] := 0.000000e+000;
   STAT28[10, 9, 5] := 0.000000e+000;
   STAT28[10, 9, 6] := 0.000000e+000;
   STAT28[10, 9, 7] := 0.000000e+000;
   STAT28[10, 9, 8] := 0.000000e+000;
   STAT28[10, 9, 9] := 0.000000e+000;
   STAT28[10, 9, 10] := 0.000000e+000;
   STAT28[10, 10, 1] := 0.000000e+000;
   STAT28[10, 10, 2] := 0.000000e+000;
   STAT28[10, 10, 3] := 0.000000e+000;
   STAT28[10, 10, 4] := 0.000000e+000;
   STAT28[10, 10, 5] := 0.000000e+000;
   STAT28[10, 10, 6] := 0.000000e+000;
   STAT28[10, 10, 7] := 0.000000e+000;
   STAT28[10, 10, 8] := 0.000000e+000;
   STAT28[10, 10, 9] := 0.000000e+000;
   STAT28[10, 10, 10] := 0.000000e+000;
   STAT29[1, 1].STAT30 := 0.000000e+000;
   STAT29[1, 1].STAT31 := 0.000000e+000;
   STAT29[1, 1].STAT32 := 0.000000e+000;
   STAT29[1, 2].STAT30 := 0.000000e+000;
   STAT29[1, 2].STAT31 := 0.000000e+000;
   STAT29[1, 2].STAT32 := 0.000000e+000;
   STAT29[1, 3].STAT30 := 0.000000e+000;
   STAT29[1, 3].STAT31 := 0.000000e+000;
   STAT29[1, 3].STAT32 := 0.000000e+000;
   STAT29[1, 4].STAT30 := 0.000000e+000;
   STAT29[1, 4].STAT31 := 0.000000e+000;
   STAT29[1, 4].STAT32 := 0.000000e+000;
   STAT29[1, 5].STAT30 := 0.000000e+000;
   STAT29[1, 5].STAT31 := 0.000000e+000;
   STAT29[1, 5].STAT32 := 0.000000e+000;
   STAT29[1, 6].STAT30 := 0.000000e+000;
   STAT29[1, 6].STAT31 := 0.000000e+000;
   STAT29[1, 6].STAT32 := 0.000000e+000;
   STAT29[1, 7].STAT30 := 0.000000e+000;
   STAT29[1, 7].STAT31 := 0.000000e+000;
   STAT29[1, 7].STAT32 := 0.000000e+000;
   STAT29[1, 8].STAT30 := 0.000000e+000;
   STAT29[1, 8].STAT31 := 0.000000e+000;
   STAT29[1, 8].STAT32 := 0.000000e+000;
   STAT29[1, 9].STAT30 := 0.000000e+000;
   STAT29[1, 9].STAT31 := 0.000000e+000;
   STAT29[1, 9].STAT32 := 0.000000e+000;
   STAT29[1, 10].STAT30 := 0.000000e+000;
   STAT29[1, 10].STAT31 := 0.000000e+000;
   STAT29[1, 10].STAT32 := 0.000000e+000;
   STAT29[2, 1].STAT30 := 0.000000e+000;
   STAT29[2, 1].STAT31 := 0.000000e+000;
   STAT29[2, 1].STAT32 := 0.000000e+000;
   STAT29[2, 2].STAT30 := 0.000000e+000;
   STAT29[2, 2].STAT31 := 0.000000e+000;
   STAT29[2, 2].STAT32 := 0.000000e+000;
   STAT29[2, 3].STAT30 := 0.000000e+000;
   STAT29[2, 3].STAT31 := 0.000000e+000;
   STAT29[2, 3].STAT32 := 0.000000e+000;
   STAT29[2, 4].STAT30 := 0.000000e+000;
   STAT29[2, 4].STAT31 := 0.000000e+000;
   STAT29[2, 4].STAT32 := 0.000000e+000;
   STAT29[2, 5].STAT30 := 0.000000e+000;
   STAT29[2, 5].STAT31 := 0.000000e+000;
   STAT29[2, 5].STAT32 := 0.000000e+000;
   STAT29[2, 6].STAT30 := 0.000000e+000;
   STAT29[2, 6].STAT31 := 0.000000e+000;
   STAT29[2, 6].STAT32 := 0.000000e+000;
   STAT29[2, 7].STAT30 := 0.000000e+000;
   STAT29[2, 7].STAT31 := 0.000000e+000;
   STAT29[2, 7].STAT32 := 0.000000e+000;
   STAT29[2, 8].STAT30 := 0.000000e+000;
   STAT29[2, 8].STAT31 := 0.000000e+000;
   STAT29[2, 8].STAT32 := 0.000000e+000;
   STAT29[2, 9].STAT30 := 0.000000e+000;
   STAT29[2, 9].STAT31 := 0.000000e+000;
   STAT29[2, 9].STAT32 := 0.000000e+000;
   STAT29[2, 10].STAT30 := 0.000000e+000;
   STAT29[2, 10].STAT31 := 0.000000e+000;
   STAT29[2, 10].STAT32 := 0.000000e+000;
   STAT29[3, 1].STAT30 := 0.000000e+000;
   STAT29[3, 1].STAT31 := 0.000000e+000;
   STAT29[3, 1].STAT32 := 0.000000e+000;
   STAT29[3, 2].STAT30 := 0.000000e+000;
   STAT29[3, 2].STAT31 := 0.000000e+000;
   STAT29[3, 2].STAT32 := 0.000000e+000;
   STAT29[3, 3].STAT30 := 0.000000e+000;
   STAT29[3, 3].STAT31 := 0.000000e+000;
   STAT29[3, 3].STAT32 := 0.000000e+000;
   STAT29[3, 4].STAT30 := 0.000000e+000;
   STAT29[3, 4].STAT31 := 0.000000e+000;
   STAT29[3, 4].STAT32 := 0.000000e+000;
   STAT29[3, 5].STAT30 := 0.000000e+000;
   STAT29[3, 5].STAT31 := 0.000000e+000;
   STAT29[3, 5].STAT32 := 0.000000e+000;
   STAT29[3, 6].STAT30 := 0.000000e+000;
   STAT29[3, 6].STAT31 := 0.000000e+000;
   STAT29[3, 6].STAT32 := 0.000000e+000;
   STAT29[3, 7].STAT30 := 0.000000e+000;
   STAT29[3, 7].STAT31 := 0.000000e+000;
   STAT29[3, 7].STAT32 := 0.000000e+000;
   STAT29[3, 8].STAT30 := 0.000000e+000;
   STAT29[3, 8].STAT31 := 0.000000e+000;
   STAT29[3, 8].STAT32 := 0.000000e+000;
   STAT29[3, 9].STAT30 := 0.000000e+000;
   STAT29[3, 9].STAT31 := 0.000000e+000;
   STAT29[3, 9].STAT32 := 0.000000e+000;
   STAT29[3, 10].STAT30 := 0.000000e+000;
   STAT29[3, 10].STAT31 := 0.000000e+000;
   STAT29[3, 10].STAT32 := 0.000000e+000;
   STAT29[4, 1].STAT30 := 0.000000e+000;
   STAT29[4, 1].STAT31 := 0.000000e+000;
   STAT29[4, 1].STAT32 := 0.000000e+000;
   STAT29[4, 2].STAT30 := 0.000000e+000;
   STAT29[4, 2].STAT31 := 0.000000e+000;
   STAT29[4, 2].STAT32 := 0.000000e+000;
   STAT29[4, 3].STAT30 := 0.000000e+000;
   STAT29[4, 3].STAT31 := 0.000000e+000;
   STAT29[4, 3].STAT32 := 0.000000e+000;
   STAT29[4, 4].STAT30 := 0.000000e+000;
   STAT29[4, 4].STAT31 := 0.000000e+000;
   STAT29[4, 4].STAT32 := 0.000000e+000;
   STAT29[4, 5].STAT30 := 0.000000e+000;
   STAT29[4, 5].STAT31 := 0.000000e+000;
   STAT29[4, 5].STAT32 := 0.000000e+000;
   STAT29[4, 6].STAT30 := 0.000000e+000;
   STAT29[4, 6].STAT31 := 0.000000e+000;
   STAT29[4, 6].STAT32 := 0.000000e+000;
